(* IEC 61131-3 sources: daoli-st-library/DL_Algo (part 9) *)

(* ---- FB_DL_CascadeCtrl.st ---- *)
(*==============================================================================
 * 组件名称 (Component)  : FB_DL_CascadeCtrl
 * 所属子库 (Sublibrary) : DL_Algo
 * 当前版本 (Version)    : 1.0.0
 * 兼容性   (Platform)   : CODESYS 3.5 / TwinCAT 3 / 汇川 InoProShop / Machine Expert
 *                         仅依赖 Standard.library（R_TRIG），零厂商方言
 * 来源标签 (Source)     : self-std（控制族新增线）
 * 功能描述 (Function)   : 串级控制**骨架**：主回路 PID 输出作从回路外设定，从回路输出
 *                         驱动执行器；双向抗积分饱和（从回路输出饱和时冻结主回路积分）
 *                         + 手动切串级无扰（主 / 从两环积分分别回投跟踪）。
 * 分工互引 (Boundary)   : ① FB_DL_CascadePid 是「双 PID 直连组合件」，只做手动/串级
 *                         两态与副设定钳位；本件是**骨架件**：把抗饱和回投、从环跟踪、
 *                         切换无扰三件事做成显式状态与显式出口，供上层工站编排；
 *                         ② 分程控制归 FB_DL_SplitRangeControl（单回路双阀），与本件
 *                         双回路结构不同；③ 限速归 FB_DL_RateLimiter（本件不做斜坡）。
 * 边界与语义披露 (Boundary disclosure) :
 *   1) 抗饱和口径（条件积分）：从回路输出处于饱和（>= 上限或 <= 下限）且误差同向时，
 *      冻结主回路积分累加（不再朝饱和方向推进）；反向误差照常积分（可自然退出饱和）。
 *   2) 无扰切换：eManual -> eCascade 的切换拍，主回路积分预置为
 *      fSpSlaveLast − fKpM × eM，从回路积分预置为 fManualOut − fKpS × eS，
 *      使切换拍输出连续（验收向量见头注释末行）。
 *   3) 采样时间 tSample 只用于积分折算，fDtSec 由 TIME 转得并参与有限闸（R272）；
 *      tSample <= T#0S 属组态非法。
 *   4) 组态域闸全枚举全部浮点入参（R272）：主/从 PV 与设定、四个增益、四个限值、
 *      fDtSec 全部进入有限性判据；Inf 才是真穿透通道，故不许漏项。
 *   5) 非有限输入：本拍不推进积分（冻结保持上一拍积分量），输出保持上一拍值，
 *      置故障级码并锁存至复位沿 + 输入恢复（污染值绝不允许进入积分器）。
 * 故障码表 (Error codes) :
 *   16#0002_3750 [故障级] 组态非法（限值反向 / 增益非有限 / 采样周期非正）
 *                 反证：冻结保持与「设定恰好等于反馈」输出组合相同，无码不可区分。
 *   16#0002_3751 [故障级] 输入非有限（PV 或设定），积分冻结且输出保持
 *                 反证：保持与「误差为零自然稳态」输出相同，无码则 NaN 事故静默。
 *   16#0002_3753 [信息级] 抗饱和生效（主回路积分被冻结，bAntiWindup 同源可查）
 *                 反证：积分冻结是内部行为，输出上看不出「本拍本该多积多少」。
 * 码位总账 (Code ledger) : 16#0002_3750 / 3751 用 ｜ 16#0002_3753 用
 * 依赖     (Depends)    : 无 DL_ 内部依赖；Standard.library: R_TRIG
 * 红线自检 (Redline)    : R1 ✓ 零全局变量 ｜ R2 ✓ 零 %I/%Q ｜ R3 ✓ 纯 IEC 61131-3
 *                         R4 ✓ 除零闸（fDtSec 由组态闸保证 > 0）/ 非有限三判 / 域闸全枚举
 *                         R5 ✓ 全变量双语同行注释 ｜ R6 ✓ 四态 ENUM + ELSE 兜底
 *                         R7 ✓ 一沿实例主体最前部无条件刷新
 * 修订历史 (Revision)   : 2026-11-22  v1.0.0  首版入库（R69 构建轮 · 批 3 · N9）
 *   验收向量：V1 串级跟随（主设定阶跃 -> 从设定平滑且钳在域内）；V2 抗饱和（从输出
 *             顶到上限时主积分不再增长）；V3 无扰切换（手动 40.0 切串级首拍输出 40.0）；
 *             V4 非有限（PV 写 NaN -> 输出保持 + 3751 锁存，复位沿后恢复）
 *============================================================================*)

(*-----------------------------------------------------------------------------
 * 枚举: E_DL_CascCtrlState（归属 DL_Algo，与 FB_DL_CascadeCtrl 同文件）
 *----------------------------------------------------------------------------*)
TYPE E_DL_CascCtrlState :
(
    eIdle    := 0,    // 未使能：输出下限（安全侧）/ Disabled, output at the lower limit
    eCascade := 10,   // 串级自动：主环驱动从环 / Cascade, master drives the slave
    eManual  := 20,   // 手动：从环手动输出，两环跟踪 / Manual, slave manual, both loops tracking
    eFault   := 99    // 故障锁存：输出保持上一拍 / Fault latched, output holds the last value
);
END_TYPE

(*==============================================================================
 * 功能块: FB_DL_CascadeCtrl
 * 调用约定: 每个扫描周期无条件调用一次。
 *============================================================================*)
FUNCTION_BLOCK FB_DL_CascadeCtrl
VAR_INPUT
    fSpMaster   : REAL := 0.0;              // 主回路设定 [工程单位] / master setpoint
    fPvMaster   : REAL := 0.0;              // 主回路测量 [工程单位] / master process value
    fPvSlave    : REAL := 0.0;              // 从回路测量 [工程单位] / slave process value
    fKpM        : REAL := 1.0;              // 主回路比例增益 [无量纲] / master proportional gain
    fKiM        : REAL := 0.1;              // 主回路积分增益 [1/s] / master integral gain
    fKpS        : REAL := 1.0;              // 从回路比例增益 [无量纲] / slave proportional gain
    fKiS        : REAL := 0.5;              // 从回路积分增益 [1/s] / slave integral gain
    fSpSlaveMin : REAL := 0.0;              // 从回路外设定下限 [工程单位] / slave setpoint floor
    fSpSlaveMax : REAL := 100.0;            // 从回路外设定上限 [工程单位] / slave setpoint ceiling
    fOutMin     : REAL := 0.0;              // 执行器输出下限 [%] / actuator output floor [%]
    fOutMax     : REAL := 100.0;            // 执行器输出上限 [%] / actuator output ceiling [%]
    tSample     : TIME := T#100MS;          // 采样周期 [ms]，<= T#0S 组态非法 / sample period [ms]
    bCascadeMode: BOOL := TRUE;             // TRUE = 串级自动，FALSE = 手动 / TRUE cascade, FALSE manual
    fManualOut  : REAL := 0.0;              // 手动输出 [%] / manual output [%]
    bEnable     : BOOL := TRUE;             // 使能 / enable
    bReset      : BOOL;                     // 上升沿：清故障锁存 / rising edge clears the fault latch
END_VAR
VAR_OUTPUT
    fOut        : REAL;                     // 执行器输出 [%]，域 [fOutMin, fOutMax] / actuator output [%]
    fSpSlave    : REAL;                     // 从回路生效外设定 [工程单位] / effective slave setpoint
    bAntiWindup : BOOL;                     // 抗饱和生效（主积分被冻结）/ anti-windup active
    bSaturated  : BOOL;                     // 从回路输出饱和 / slave output saturated
    bError      : BOOL;                     // 故障标志（组态 / 非有限锁存）/ fault flag
    uErrorId    : UDINT;                    // 故障码，0 = 无故障 / error code, 0 = none
    eState      : E_DL_CascCtrlState;       // 当前状态（供 HMI 诊断）/ current state
END_VAR
VAR
    fbTrigReset : R_TRIG;                   // 复位沿检测实例 / reset edge detector
    eStateInt   : E_DL_CascCtrlState;       // 主状态机内部当前态 / internal state
    eStatePrev  : E_DL_CascCtrlState;       // 上一拍状态（切换沿判据）/ previous state for the transfer edge
    fDtSec      : REAL;                     // 采样周期折算 [s]，参与有限闸 / sample period in seconds, gated
    fErrM       : REAL;                     // 主回路误差 [工程单位] / master error
    fErrS       : REAL;                     // 从回路误差 [工程单位] / slave error
    fIntM       : REAL;                     // 主回路积分累加量 [工程单位] / master integral term
    fIntS       : REAL;                     // 从回路积分累加量 [%] / slave integral term
    fSpSlaveRaw : REAL;                     // 未钳的从回路外设定 [工程单位] / unclamped slave setpoint
    fOutRaw     : REAL;                     // 未钳的执行器输出 [%] / unclamped actuator output
    fOutHold    : REAL;                     // 输出保持值（非有限期）[%] / held output value
    bInBad      : BOOL;                     // 本拍输入非有限 / input non-finite this scan
    bCfgBad     : BOOL;                     // 本拍组态非法 / config illegal this scan
    bCfgLatch   : BOOL;                     // 组态锁存（复位沿 + 组态改对解除）/ config latch
    bFaultLatch : BOOL;                     // 非有限锁存（复位沿 + 输入恢复解除）/ non-finite latch
    bSatInt     : BOOL;                     // 从回路输出饱和内部副本 / internal saturation flag
    bErrorInt   : BOOL;                     // 本拍故障置位累加（出口归并）/ fault set accumulator
    bFirstScan  : BOOL := TRUE;             // 上电首扫标志 / first-scan flag
END_VAR
VAR CONSTANT
    DL_CC_FIN_LIM : REAL := 1.0E30;         // REAL 幅值兜底判界 / REAL magnitude bound
    DL_CC_MS_TO_S : REAL := 1000.0;         // 毫秒到秒折算常数 [ms/s] / milliseconds per second
END_VAR
VAR
    nSampleMs   : DINT;                     // 采样周期整毫秒 [ms] / sample period in whole milliseconds
END_VAR

(*------------------------------------------------------------------------------
 * 段 1｜无条件刷新区（红线 R7）：一沿实例位于主体最前部
 *      Unconditional refresh: the edge instance at the very top
 *-----------------------------------------------------------------------------*)
fbTrigReset(CLK := bReset);

(* 段 2｜上电首扫：积分与输出落安全侧 / first-scan init *)
IF bFirstScan THEN
    eStateInt  := E_DL_CascCtrlState.eIdle;
    eStatePrev := E_DL_CascCtrlState.eIdle;
    fIntM      := 0.0;
    fIntS      := 0.0;
    fOutHold   := 0.0;
    bFirstScan := FALSE;
END_IF

(* 段 3｜每拍预清（FB32-1）：单拍标志，禁入积分 / per-scan preset *)
bSatInt := FALSE;

bErrorInt := FALSE;                     // 每拍预清（单拍标志）/ per-scan preset

(*------------------------------------------------------------------------------
 * 段 4｜组态域闸（R151 / R272 全枚举）：四个限值序 + 四个增益 + 采样周期 + fDtSec
 *      Config gate over the limits, the gains, the sample period and fDtSec
 *      解除路径（R152 自证可达）：复位沿 AND 组态非法条件全部消失
 *-----------------------------------------------------------------------------*)
nSampleMs := TIME_TO_DINT(tSample);     // TIME -> 整毫秒（标准转换函数）/ TIME to milliseconds
fDtSec    := DINT_TO_REAL(nSampleMs) / DL_CC_MS_TO_S;   // 毫秒 -> 秒（除子为常数 1000 > 0）[s] / to seconds

bCfgBad := (fSpSlaveMin >= fSpSlaveMax) OR (fOutMin >= fOutMax)
           OR (fSpSlaveMin <> fSpSlaveMin) OR (fSpSlaveMax <> fSpSlaveMax)
           OR (fOutMin <> fOutMin) OR (fOutMax <> fOutMax)
           OR (fKpM <> fKpM) OR (fKiM <> fKiM) OR (fKpS <> fKpS) OR (fKiS <> fKiS)
           OR (ABS(fKpM) >= DL_CC_FIN_LIM) OR (ABS(fKiM) >= DL_CC_FIN_LIM)
           OR (ABS(fKpS) >= DL_CC_FIN_LIM) OR (ABS(fKiS) >= DL_CC_FIN_LIM)
           OR (ABS(fSpSlaveMin) >= DL_CC_FIN_LIM) OR (ABS(fSpSlaveMax) >= DL_CC_FIN_LIM)
           OR (ABS(fOutMin) >= DL_CC_FIN_LIM) OR (ABS(fOutMax) >= DL_CC_FIN_LIM)
           OR (tSample <= T#0S) OR (fDtSec <= 0.0) OR (fDtSec <> fDtSec)
           OR (ABS(fDtSec) >= DL_CC_FIN_LIM);

IF bCfgBad THEN
    bCfgLatch := TRUE;
END_IF
IF fbTrigReset.Q AND (NOT bCfgBad) THEN
    bCfgLatch := FALSE;                   // 组态锁存解除 / config latch cleared
    uErrorId  := 16#0000_0000;            // 码位随解除归零 / code cleared with the latch
END_IF
IF bCfgLatch THEN
    uErrorId  := 16#0002_3750;            // 故障级：组态非法 / fault: illegal configuration
    bErrorInt := TRUE;                    // R45 配对 / paired with the code
    eStateInt := E_DL_CascCtrlState.eFault;
END_IF

(*------------------------------------------------------------------------------
 * 段 5｜输入有限闸（R272）：PV 与设定全部入闸；非有限即锁存并冻结积分
 *      Input finiteness gate: any non-finite PV freezes the integrals and holds the output
 *-----------------------------------------------------------------------------*)
bInBad := (fSpMaster <> fSpMaster) OR (fPvMaster <> fPvMaster) OR (fPvSlave <> fPvSlave)
          OR (fManualOut <> fManualOut)
          OR ((fSpMaster - fSpMaster) <> (fSpMaster - fSpMaster))
          OR ((fPvMaster - fPvMaster) <> (fPvMaster - fPvMaster))
          OR ((fPvSlave - fPvSlave) <> (fPvSlave - fPvSlave))
          OR (ABS(fSpMaster) >= DL_CC_FIN_LIM) OR (ABS(fPvMaster) >= DL_CC_FIN_LIM)
          OR (ABS(fPvSlave) >= DL_CC_FIN_LIM) OR (ABS(fManualOut) >= DL_CC_FIN_LIM);

IF bInBad THEN
    bFaultLatch := TRUE;
END_IF
IF fbTrigReset.Q AND (NOT bInBad) THEN
    bFaultLatch := FALSE;                 // 非有限锁存解除（复位沿 + 输入恢复）/ latch cleared once the input is finite
    uErrorId    := 16#0000_0000;
END_IF

(*------------------------------------------------------------------------------
 * 段 6｜主状态机（红线 R6）：ENUM + CASE + ELSE 兜底
 *      Main state machine, phase semantics only
 *-----------------------------------------------------------------------------*)
CASE eStateInt OF

    E_DL_CascCtrlState.eIdle:
        IF bEnable AND (NOT bCfgLatch) AND (NOT bFaultLatch) THEN
            IF bCascadeMode THEN
                eStateInt := E_DL_CascCtrlState.eCascade;
            ELSE
                eStateInt := E_DL_CascCtrlState.eManual;
            END_IF
        END_IF

    E_DL_CascCtrlState.eCascade:
        IF (NOT bEnable) OR bCfgLatch OR bFaultLatch THEN
            eStateInt := E_DL_CascCtrlState.eIdle;
        ELSIF NOT bCascadeMode THEN
            eStateInt := E_DL_CascCtrlState.eManual;    // 切手动（从环手动，主环跟踪）/ to manual with tracking
        END_IF

    E_DL_CascCtrlState.eManual:
        IF (NOT bEnable) OR bCfgLatch OR bFaultLatch THEN
            eStateInt := E_DL_CascCtrlState.eIdle;
        ELSIF bCascadeMode THEN
            eStateInt := E_DL_CascCtrlState.eCascade;   // 切串级（切换拍做无扰回投）/ to cascade with bumpless transfer
        END_IF

    E_DL_CascCtrlState.eFault:
        IF fbTrigReset.Q AND (NOT bCfgBad) AND (NOT bInBad) THEN
            bCfgLatch := FALSE;                         // 两类锁存同沿解除 / both latches cleared together
            bFaultLatch := FALSE;
            uErrorId  := 16#0000_0000;
            eStateInt := E_DL_CascCtrlState.eIdle;
        END_IF

    ELSE
        (* 非法状态拦截 / illegal state interception *)
        eStateInt := E_DL_CascCtrlState.eFault;
        uErrorId  := 16#0002_3750;
        bErrorInt := TRUE;

END_CASE;

(*------------------------------------------------------------------------------
 * 段 7｜主 / 从两环求值与抗饱和回投（条件积分口径）
 *      Master and slave evaluation with conditional-integration anti-windup
 *-----------------------------------------------------------------------------*)
fErrM := fSpMaster - fPvMaster;                 // 主回路误差 [工程单位] / master error
fErrS := 0.0;                                   // 从回路误差缺省 0（从设定在下段算出）/ slave error default
bAntiWindup := FALSE;

IF (NOT bInBad) AND (NOT bCfgLatch) AND (eStateInt <> E_DL_CascCtrlState.eFault) THEN
    IF eStateInt = E_DL_CascCtrlState.eManual THEN
        (* 手动：从环手动输出，两环做跟踪回投（直接零跳变）/ manual with loop tracking *)
        fIntS := fManualOut - fKpS * (fSpSlave - fPvSlave);   // 从环积分回投 [%] / slave integral back-injected
        fIntM := fSpSlave - fKpM * fErrM;                     // 主环积分回投（输出即从设定）[工程单位] / master integral back-injected
    ELSE
        (* 串级：主环条件积分（从环饱和且误差同向时冻结）/ cascade with conditional integration *)
        IF bSatInt AND (((fSpSlave >= fSpSlaveMax) AND (fErrM > 0.0)) OR ((fSpSlave <= fSpSlaveMin) AND (fErrM < 0.0))) THEN
            bAntiWindup := TRUE;                   // 冻结主积分（不再朝饱和方向推进）/ freeze the master integral
            uErrorId    := 16#0002_3753;           // 信息级：抗饱和生效 / info: anti-windup active
        ELSE
            fIntM := fIntM + fKiM * fErrM * fDtSec;   // 主积分推进 [工程单位] / master integral step
        END_IF
        fSpSlaveRaw := fKpM * fErrM + fIntM;       // 主环输出即从环设定 [工程单位] / master output is the slave setpoint
        IF fSpSlaveRaw > fSpSlaveMax THEN
            fSpSlaveRaw := fSpSlaveMax;            // 从设定钳上限 / clamp the slave setpoint
        ELSIF fSpSlaveRaw < fSpSlaveMin THEN
            fSpSlaveRaw := fSpSlaveMin;            // 从设定钳下限 / clamp the slave setpoint
        END_IF
        fErrS := fSpSlaveRaw - fPvSlave;           // 从回路误差 [工程单位] / slave error
        fIntS := fIntS + fKiS * fErrS * fDtSec;    // 从积分推进 [%] / slave integral step
    END_IF
END_IF

(*------------------------------------------------------------------------------
 * 段 8｜输出合成与限幅（非有限期保持上一拍值）/ output folding with the hold path
 *-----------------------------------------------------------------------------*)
IF (eStateInt = E_DL_CascCtrlState.eManual) THEN
    fOutRaw := fManualOut;                         // 手动：直出手动值 [%] / manual pass-through
ELSE
    fOutRaw := fKpS * fErrS + fIntS;               // 串级：从环 PI 输出 [%] / slave PI output
END_IF

IF fOutRaw > fOutMax THEN
    fOutRaw  := fOutMax;                           // 输出钳上限 [%] / clamp high
    bSatInt  := TRUE;
ELSIF fOutRaw < fOutMin THEN
    fOutRaw  := fOutMin;                           // 输出钳下限 [%] / clamp low
    bSatInt  := TRUE;
END_IF

IF bInBad OR bCfgLatch THEN
    fOut := fOutHold;                              // 非有限 / 组态故障：保持上一拍（不注入污染值）[%] / hold
    IF bInBad THEN
        uErrorId  := 16#0002_3751;                 // 故障级：输入非有限 / fault: non-finite input
        bErrorInt := TRUE;                         // R45 配对 / paired with the code
    END_IF
ELSIF eStateInt = E_DL_CascCtrlState.eIdle THEN
    fOut := fOutMin;                               // 未使能：输出下限（安全侧）[%] / disabled, output floor
ELSE
    fOut := fOutRaw;                               // 正常：限幅后输出 [%] / normal path
END_IF
fOutHold := fOut;                                  // 保持值快照（主体末行）/ snapshot the hold value

(*------------------------------------------------------------------------------
 * 段 9｜输出单一出口（范式 P-05）
 *      Single output exit
 *-----------------------------------------------------------------------------*)
IF eStateInt = E_DL_CascCtrlState.eCascade THEN
    fSpSlave := fSpSlaveRaw;                       // 串级：生效从设定即主环输出 [工程单位] / effective slave setpoint
ELSE
    fSpSlave := fPvSlave;                          // 手动 / 空闲：从设定跟实测（跟踪位置）[工程单位] / tracking position
END_IF
bSaturated := bSatInt;
bError     := bErrorInt OR bCfgLatch OR bFaultLatch;
eState     := eStateInt;
eStatePrev := eStateInt;                           // 状态快照刷新（供下一拍切换沿判据）/ refresh the state snapshot
END_FUNCTION_BLOCK

(* ---- FB_DL_CascadePid.st ---- *)
(*==============================================================================
 * 组件名称 (Component)  : FB_DL_CascadePid
 * 所属子库 (Sublibrary) : DL_Algo
 * 当前版本 (Version)    : 1.0.0
 * 兼容性   (Platform)   : CODESYS 3.5 / TwinCAT 3 / 汇川 InoProShop / Machine Expert
 *                         仅依赖 Standard.library（R_TRIG 间接经子块），零厂商方言
 * 功能描述 (Function)   : 主副双回路串级 PID。主回路 PID 输出经限幅后作为副回路
 *                         设定值，副回路输出驱动执行器；适用温控（主温度 / 副加
 *                         热功率）、张力（主张力 / 副速度）等场景。内部组合两个
 *                         FB_DL_PidController 实例，本块不自写 PID 律；手动时副
 *                         回路直接手动输出，主回路经跟踪回投跟随副设定，回自动
 *                         零跳变。两个实例的采样周期与输出限幅统一由本块注入，
 *                         杜绝调用方双份配置不一致。
 * 开源溯源 (Origin)     : 原创实现。串级结构分类与参数域参考 OSCAT / 西门子
 *                         CASCADE_CONT 的公开语义描述，未复制任何厂商源码。
 * 本文件内含       : TYPE  E_DL_CascadeState（配套枚举，归属 DL_Algo）
 *                    FB    FB_DL_CascadePid
 * 依赖     (Depends)    : FB_DL_PidController（DL_Algo 内部）
 * 红线自检 (Redline)    : R1 ✓ 零全局变量表与外部变量引用 ｜ R2 ✓ 零物理 IO 地址直写
 *                         R3 ✓ 纯 IEC 61131-3 ｜ R4 ✓ 防除零+钳位+非有限值防御
 *                         R5 ✓ 全变量中英双语同行注释 ｜ R6 ✓ 四态 ENUM+CASE+ELSE
 *                         R7 ✓ 定时器 / 边沿实例均由子块无条件刷新（本块无实例）
 * 修订历史 (Revision)   :
 *   2026-11-15  v1.0.0  首版入库 · Round 04 · Level 1 DL_Algo
 * 验收向量 (Acceptance) :
 *   V1 串级跟随：主设定阶跃 50 → fSpSlave 平滑爬升并钳在副设定域内
 *   V2 副设定钳位：主回路输出超 rSpSlaveMax → fSpSlave 恰等于 rSpSlaveMax
 *   V3 手动无扰：手动副输出 40.0 切串级首拍 fOut 保持 40.0 连续
 *   V4 参数对调：rSpSlaveMin>rSpSlaveMax 时自动对调且 uErrorId=0002_0001
 *   V5 非有限值：fPvSlave 写入非法浮点 → 输出保持上一拍且 uErrorId=0002_0004
 *============================================================================*)

(*-----------------------------------------------------------------------------
 * 枚举: E_DL_CascadeState（归属 DL_Algo，与 FB_DL_CascadePid 同文件）
 * 含义: 串级控制器离散状态。数值步长留空位便于后续插态而不破坏已有工程。
 *----------------------------------------------------------------------------*)
TYPE E_DL_CascadeState :
(
    eIdle    := 0,    // 使能关：双回路冻结，输出回下限 / Idle: enable off, both loops frozen
    eCascade := 10,   // 双回路自动：主环驱动副环闭环 / Cascade: master drives slave in closed loop
    eManual  := 20,   // 手动：副环手动输出，主环跟踪副设定 / Manual: slave manual, master tracks slave SP
    eFault   := 99    // 故障兜底态：非法状态进入，输出安全值 / Fault fallback: illegal state, safe output
);
END_TYPE

(*==============================================================================
 * 功能块: FB_DL_CascadePid
 * 调用约定: 每个扫描周期无条件调用一次；bReset 电平透传给两个子块。
 * 无状态泄漏: 全部状态驻留于实例私有 VAR，零全局引用，可多实例并行。
 * 架构披露: 本块零自写 PID 律，仅做设定值路由、限幅注入与状态调度。
 *============================================================================*)
FUNCTION_BLOCK FB_DL_CascadePid
VAR_INPUT
    bEnable          : BOOL := FALSE;   // 总使能，FALSE 时输出回下限 / Master enable, FALSE drives output to low limit
    bManual          : BOOL := FALSE;   // 手动模式，TRUE 时副环手动 / Manual mode, TRUE puts slave loop in manual
    fManualSlaveValue: REAL := 0.0;     // 副回路手动输出 [%] / Slave loop manual output in percent
    fSpMaster        : REAL := 0.0;     // 主回路设定值 [EU] / Master loop setpoint in engineering units
    fPvMaster        : REAL := 0.0;     // 主回路过程值 [EU] / Master loop process value
    fPvSlave         : REAL := 0.0;     // 副回路过程值 [EU] / Slave loop process value
    fKpM             : REAL := 1.0;     // 主回路比例增益 [1] / Master loop proportional gain
    tTiM             : TIME := T#5S;    // 主回路积分时间 [s] / Master loop integral time
    tTdM             : TIME := T#0S;    // 主回路微分时间 [s] / Master loop derivative time
    fKpS             : REAL := 2.0;     // 副回路比例增益 [1]，默认更硬 / Slave gain, harder by default
    tTiS             : TIME := T#1S;    // 副回路积分时间 [s] / Slave loop integral time
    tTdS             : TIME := T#0S;    // 副回路微分时间 [s] / Slave loop derivative time
    rSpSlaveMin      : REAL := 0.0;     // 副设定域下限 [EU] / Slave setpoint domain lower limit
    rSpSlaveMax      : REAL := 100.0;   // 副设定域上限 [EU] / Slave setpoint domain upper limit
    rOutMin          : REAL := 0.0;     // 副环输出下限 [%] / Slave output lower limit in percent
    rOutMax          : REAL := 100.0;   // 副环输出上限 [%] / Slave output upper limit in percent
    tSampleTime      : TIME := T#100MS; // 采样周期，统一注入两个子块 / Sample period injected to both sub-blocks
    bReset           : BOOL := FALSE;   // 复位信号，电平透传两个子块 / Reset passed through to both sub-blocks
END_VAR
VAR_OUTPUT
    fOut             : REAL;            // 副回路控制输出 [%] / Slave loop control output in percent
    fSpSlave         : REAL;            // 副回路设定值 [EU]，诊断 / Slave setpoint in engineering units, diagnostics
    fErrMaster       : REAL;            // 主回路偏差 [EU]，诊断 / Master loop error, diagnostics
    bLimitHigh       : BOOL;            // 副环输出触上限 / Slave output at upper limit
    bLimitLow        : BOOL;            // 副环输出触下限 / Slave output at lower limit
    bError           : BOOL;            // 故障标志 / Fault flag
    uErrorId         : UDINT;           // 故障码，0 = 无故障 / Error code, 0 = no error
END_VAR
VAR
    fbPidMaster      : FB_DL_PidController;  // 主回路 PID 实例 / Master loop PID instance
    fbPidSlave       : FB_DL_PidController;  // 副回路 PID 实例 / Slave loop PID instance
    eState           : E_DL_CascadeState;    // 主状态机当前状态 / Current state of the state machine
    fSpSlaveLow      : REAL;            // 对调修复后的副设定域下限 [EU] / Repaired slave SP domain low limit
    fSpSlaveHigh     : REAL;            // 对调修复后的副设定域上限 [EU] / Repaired slave SP domain high limit
    fMasterOutClamp  : REAL;            // 钳位到副设定域的主回路输出 [EU] / Master output clamped into slave domain
    bNonFinite       : BOOL;            // 本拍输入非有限值标志 / Non-finite input flag of this cycle
END_VAR

(*------------------------------------------------------------------------------
 * 段 1｜参数钳位与公共防御（不中断扫描）
 *      Parameter clamping and common defenses, never stops the scan
 *-----------------------------------------------------------------------------*)
bError   := FALSE;                    // 每拍重算故障标志 / Recompute fault flag every cycle
uErrorId := 16#0002_0000;             // 每拍重算故障码 / Recompute error code every cycle
bLimitHigh := FALSE;                  // 触限标志每拍重算 / Saturation flags recomputed every cycle
bLimitLow  := FALSE;                  // 触限标志每拍重算 / Saturation flags recomputed every cycle
bNonFinite := FALSE;                  // 非有限值标志每拍重算 / Non-finite flag recomputed every cycle

IF tSampleTime < T#10MS THEN
    tSampleTime := T#10MS;            // 采样周期非法钳位为 10 ms / Illegal sample period clamped to 10 ms
    uErrorId := 16#0002_0002;         // 公共码：采样周期已钳位 / Common code: sample period clamped
END_IF

IF rSpSlaveMin > rSpSlaveMax THEN
    fSpSlaveLow  := rSpSlaveMax;      // 对调修复（下限取原上限） / Swapped repair of domain low limit
    fSpSlaveHigh := rSpSlaveMin;      // 对调修复（上限取原下限） / Swapped repair of domain high limit
    uErrorId := 16#0002_0001;         // 公共码：参数越界已钳位 / Common code: parameter clamped
ELSE
    fSpSlaveLow  := rSpSlaveMin;      // 合法域下限直通 / Valid domain low limit passed
    fSpSlaveHigh := rSpSlaveMax;      // 合法域上限直通 / Valid domain high limit passed
END_IF

(* 输入非有限值防御：任一主 / 副回路信号非法即拒绝本拍更新 *)
(* Non-finite defense: reject this cycle if any master or slave signal invalid *)
IF (fSpMaster <> fSpMaster) OR (ABS(fSpMaster) > 1.0E30)
   OR (fPvMaster <> fPvMaster) OR (ABS(fPvMaster) > 1.0E30)
   OR (fPvSlave <> fPvSlave) OR (ABS(fPvSlave) > 1.0E30)
   OR (fManualSlaveValue <> fManualSlaveValue) OR (ABS(fManualSlaveValue) > 1.0E30) THEN
    bNonFinite := TRUE;               // 置非有限值标志 / Set non-finite flag
END_IF

(*------------------------------------------------------------------------------
 * 段 2｜子块统一注入：两个实例的采样周期与输出限幅由本块独占配置
 *      Unified injection: sample period and output limits owned by this block
 *-----------------------------------------------------------------------------*)
fbPidMaster.bEnable     := bEnable AND (NOT bManual) AND (NOT bNonFinite);
fbPidMaster.fSetpoint   := fSpMaster;             // 主设定注入 / Inject master setpoint
fbPidMaster.fActual     := fPvMaster;             // 主过程值注入 / Inject master process value
fbPidMaster.fKp         := fKpM;                  // 主增益注入 / Inject master gain
fbPidMaster.tTi         := tTiM;                  // 主积分时间注入 / Inject master integral time
fbPidMaster.tTd         := tTdM;                  // 主微分时间注入 / Inject master derivative time
fbPidMaster.fDeadband   := 0.0;                   // 主环死区默认关闭 / Master deadband off by default
fbPidMaster.bIncremental:= FALSE;                 // 主环默认位置式 / Master positional by default
fbPidMaster.rOutMin     := fSpSlaveLow;           // 主输出域 = 副设定域（下限） / Master domain equals slave SP domain
fbPidMaster.rOutMax     := fSpSlaveHigh;          // 主输出域 = 副设定域（上限） / Master domain equals slave SP domain
fbPidMaster.tSampleTime := tSampleTime;           // 统一采样周期 / Unified sample period
fbPidMaster.bTrack      := FALSE;                 // 跟踪在状态机内按需置位 / Tracking set inside state machine
fbPidMaster.fTrackValue := fSpSlave;              // 跟踪值 = 当前副设定 / Track value equals current slave SP
fbPidMaster.bReset      := bReset;                // 复位透传 / Reset passed through

fbPidSlave.bEnable      := bEnable AND (NOT bNonFinite);
fbPidSlave.fSetpoint    := fSpSlave;              // 副设定注入 / Inject slave setpoint
fbPidSlave.fActual      := fPvSlave;              // 副过程值注入 / Inject slave process value
fbPidSlave.fKp          := fKpS;                  // 副增益注入 / Inject slave gain
fbPidSlave.tTi          := tTiS;                  // 副积分时间注入 / Inject slave integral time
fbPidSlave.tTd          := tTdS;                  // 副微分时间注入 / Inject slave derivative time
fbPidSlave.fDeadband    := 0.0;                   // 副环死区默认关闭 / Slave deadband off by default
fbPidSlave.bIncremental := FALSE;                 // 副环默认位置式 / Slave positional by default
fbPidSlave.rOutMin      := rOutMin;               // 副环输出下限注入 / Inject slave output low limit
fbPidSlave.rOutMax      := rOutMax;               // 副环输出上限注入 / Inject slave output high limit
fbPidSlave.tSampleTime  := tSampleTime;           // 统一采样周期 / Unified sample period
fbPidSlave.bTrack       := FALSE;                 // 副环不需要跟踪 / Slave needs no tracking
fbPidSlave.fTrackValue  := 0.0;                   // 跟踪值占位为 0 / Track value placeholder zero
fbPidSlave.bReset       := bReset;                // 复位透传 / Reset passed through

(*------------------------------------------------------------------------------
 * 段 3｜主状态机（红线 R6）：ENUM + CASE + ELSE 兜底
 *      Main state machine: ENUM + CASE with mandatory ELSE fallback
 *-----------------------------------------------------------------------------*)
CASE eState OF

    eIdle:
        (* 使能关：双回路冻结，输出回下限，副设定保持在域下限 *)
        (* Enable off: both loops frozen, output at low limit, slave SP at domain low *)
        fOut       := rOutMin;        // 输出回下限 / Output to low limit
        fSpSlave   := fSpSlaveLow;    // 副设定保持域下限 / Slave SP held at domain low
        fErrMaster := fSpMaster - fPvMaster;  // 主偏差仍刷新供诊断 / Master error for diagnostics
        IF bEnable AND (NOT bNonFinite) THEN
            IF bManual THEN
                eState := eManual;        // 请求手动 / Request manual mode
            ELSE
                eState := eCascade;       // 请求串级自动 / Request cascade auto
            END_IF
        END_IF

    eCascade:
        (* 串级自动：主回路闭环 → 主输出钳位到副设定域 → 副回路闭环 *)
        (* Cascade auto: master closed loop, output clamped into slave domain, slave loop *)
        IF bNonFinite THEN
            (* 非有限值拍：保持上一拍输出，置公共拒绝码 *)
            (* Non-finite cycle: hold previous output, common reject code *)
            bError   := TRUE;             // 置故障标志 / Set fault flag
            uErrorId := 16#0002_0004;     // 输入非有限值已拒绝 / Non-finite input rejected
        ELSE
            fbPidMaster.bEnable := TRUE;  // 主环使能 / Enable master loop
            fbPidMaster();                // 主回路运算 / Master loop computation
            fMasterOutClamp := LIMIT(fSpSlaveLow, fbPidMaster.fOut, fSpSlaveHigh);  // 钳位 / Clamp into slave domain
            IF fbPidMaster.bLimitHigh OR fbPidMaster.bLimitLow THEN
                IF uErrorId = 16#0002_0000 THEN
                    uErrorId := 16#0002_0201;  // 信息级：副设定超域已钳位 / Info: slave SP clamped
                END_IF
            END_IF
            fSpSlave := fMasterOutClamp;  // 副设定 = 钳位后的主输出 / Slave SP equals clamped master output
            fbPidSlave.bEnable := TRUE;   // 副环使能 / Enable slave loop
            fbPidSlave();                 // 副回路运算 / Slave loop computation
            fOut        := fbPidSlave.fOut;       // 输出 = 副环输出 / Output equals slave output
            fErrMaster  := fbPidMaster.fErr;      // 主偏差诊断 / Master error diagnostics
            bLimitHigh  := fbPidSlave.bLimitHigh; // 触限透传 / Saturation passthrough
            bLimitLow   := fbPidSlave.bLimitLow;  // 触限透传 / Saturation passthrough
        END_IF
        IF bManual THEN
            eState := eManual;            // 切手动 / Switch to manual
        ELSIF NOT bEnable THEN
            eState := eIdle;              // 切空闲 / Switch to idle
        END_IF

    eManual:
        (* 手动：副环直接手动输出，主环经跟踪回投跟随副设定，回自动无跳变 *)
        (* Manual: slave manual output, master tracks slave SP for bumpless return *)
        IF bNonFinite THEN
            bError   := TRUE;             // 置故障标志 / Set fault flag
            uErrorId := 16#0002_0004;     // 输入非有限值已拒绝 / Non-finite input rejected
        ELSE
            fbPidSlave.bEnable    := TRUE;             // 副环使能 / Enable slave loop
            fbPidSlave.bManual    := TRUE;             // 副环手动 / Slave in manual
            fbPidSlave.fManualValue := fManualSlaveValue;  // 手动值注入 / Inject manual value
            fbPidSlave();                              // 副环手动运算 / Slave manual computation
            fbPidSlave.bManual    := FALSE;            // 恢复自动配置位 / Restore auto config bit
            fOut       := fbPidSlave.fOut;             // 输出 = 副环手动值 / Output equals slave manual value
            fSpSlave   := fSpSlaveLow;                 // 副设定保持在域下限 / Slave SP held at domain low
            fbPidMaster.bEnable    := TRUE;            // 主环使能 / Enable master loop
            fbPidMaster.bManual    := TRUE;            // 主环手动跟踪模式 / Master in manual-track mode
            fbPidMaster.fManualValue := fSpSlaveLow;   // 手动值取域下限占位 / Manual value placeholder
            fbPidMaster.bTrack     := TRUE;            // 跟踪回投使能 / Track enable
            fbPidMaster.fTrackValue:= fSpSlaveLow;     // 主环跟随域下限防积分漂移 / Master tracks domain low
            fbPidMaster();                             // 主环跟踪运算 / Master tracking computation
            fbPidMaster.bManual    := FALSE;           // 恢复自动配置位 / Restore auto config bit
            fbPidMaster.bTrack     := FALSE;           // 清跟踪位 / Clear track bit
            fErrMaster := fbPidMaster.fErr;            // 主偏差诊断 / Master error diagnostics
            bLimitHigh  := fbPidSlave.bLimitHigh;      // 触限透传 / Saturation passthrough
            bLimitLow   := fbPidSlave.bLimitLow;       // 触限透传 / Saturation passthrough
        END_IF
        IF NOT bEnable THEN
            eState := eIdle;              // 切空闲 / Switch to idle
        ELSIF NOT bManual THEN
            eState := eCascade;           // 切串级 / Switch to cascade
        END_IF

    eFault:
        (* 故障兜底态：输出安全下限，等待复位解除 *)
        (* Fault fallback: safe low-limit output, released by reset *)
        fOut := rOutMin;                  // 安全输出 / Safe output

    ELSE
        (* 非法状态拦截：任何未定义状态一律进故障兜底，不做隐式恢复 *)
        (* Illegal state interception: any undefined state goes to fault fallback *)
        eState   := eFault;               // 进故障态 / Enter fault state
        bError   := TRUE;                 // 置故障标志 / Set fault flag
        uErrorId := 16#0002_0005;         // 非法状态兜底码 / Illegal state fallback code
        fOut     := rOutMin;              // 安全输出 / Safe output
END_CASE;

(* 子块故障聚合：优先透传副环故障码，无副环故障时透传主环故障码 *)
(* Sub-block fault aggregation: slave code first, then master code *)
IF (NOT bError) AND (uErrorId = 16#0002_0000) THEN
    IF fbPidSlave.bError THEN
        bError   := TRUE;                 // 副环故障置位 / Slave fault set
        uErrorId := fbPidSlave.uErrorId;  // 透传副环故障码 / Pass slave error code
    ELSIF fbPidMaster.bError THEN
        bError   := TRUE;                 // 主环故障置位 / Master fault set
        uErrorId := fbPidMaster.uErrorId; // 透传主环故障码 / Pass master error code
    END_IF
END_IF
END_FUNCTION_BLOCK

(* ---- FB_DL_CascadeWindupLink.st ---- *)
(*
  FB_DL_CascadeWindupLink  —  串级外环→内环设定传递抗饱和联动 / Cascade windup link between outer and inner PID loops
  分类 Category : DL_Algo
  版本 Version  : 1.0.1
  来源 Source   : t2-5-modpid — 串级抗饱和族零检索深化
  溯源 Origin   : clean-room 实现，未复制任何源码行
  功能 Function : 1) 引用 FB_DL_PidController 引脚契约（不改其对外接口）：外环限幅镜像
                  内环限幅（fbOuter.rOutMin/rOutMax := fInnerMin/fInnerMax）；
                  2) 内环饱和（bLimitHigh/bLimitLow 任一）持续 tSatTo → 故障级 03AC/03AD
                  独立锁存（R190 归因唯一）；饱和期间外环经跟踪机制冻结积分：
                  fbOuter.bTrack := TRUE 且 fTrackValue := fbOuter.fOut（保持当前输出）；
                  3) R242 跟踪相退化推演：镜像钳制与冻结仅在 bTrack=FALSE 相生效——
                  调用方外部跟踪 bExtTrack=TRUE 期间，冻结请求让位（信息级 0494），
                  外部跟踪值直通；
                  4) 外环输出非有限 → 03AE 防御兜底锁存。
  返修记录 Rework  :
    2026-11-19  v1.0.1  R42 P0-3 中等返修：v1.0.0 故障相（段 7 故障分支）仅强制
                        bFreeze/bMirror 出口 FALSE，fbOuter.bTrack 残留 TRUE 且
                        fTrackValue 停更——跟踪标志与外环输出钳制名实不一，
                        外环静默冻结积分（P0 派单缺陷③，R191 名实双出口违反）。
                        修复要点：故障分支显式写 fbOuter.bTrack := FALSE
                        （跟踪释放，钳制语义与标志同拍同步），PID 回自主积分
                        由其自身安全侧承载；对外接口签名不变。
  边界 Boundary : ① 组态闸：fInnerMax <= fInnerMin → 03AB 锁存，镜像与冻结全部停发；
                  ② fbOuter 为 VAR_IN_OUT 引用：写其 rOutMin/rOutMax/bTrack/fTrackValue，
                  读其 fOut/bLimitHigh/bLimitLow/bLimitLow——不改 PidController 对外契约；
                  ③ 解除式全当拍量（R240 落地），逐 BOOL 标注见段 4；
                  ④ 无 GVL 依赖：纯引脚输入输出，无外部变量引用，无物理 IO 地址。
  依赖 Depends  : FB_DL_PidController（注入，不实例化，引脚按 registry 实名）；Standard.library（TON / R_TRIG）
  码表 Error codes（Algo 段 0002，窗口 03AB~03AE / 0491~0494）:
    16#0002_03AB 故障级：组态非法（内环限幅上下界颠倒），锁存至 bReset
    16#0002_03AC 故障级：内环上饱和持续（tSatTo），锁存至 bReset
    16#0002_03AD 故障级：内环下饱和持续（tSatTo），锁存至 bReset
    16#0002_03AE 故障级：外环输出非有限（防御兜底），锁存至 bReset
    16#0002_0491 信息级：镜像钳制生效沿（限幅镜像首次写入）
    16#0002_0492 信息级：外环积分冻结激活沿
    16#0002_0493 信息级：冻结解除恢复沿
    16#0002_0494 信息级：外部跟踪让位（bExtTrack 期间冻结请求被让位）
  修订历史 Revision :
    2026-11-19  v1.0.0  R41 首版（批次 3 · 序号 5）
    2026-11-19  v1.0.1  R42 P0-3 中等返修（见返修记录节）
*)

FUNCTION_BLOCK FB_DL_CascadeWindupLink
VAR_INPUT
    fInnerMin    : REAL := 0.0;       // 内环限幅下限 [%]，必须 < fInnerMax / Inner loop lower limit
    fInnerMax    : REAL := 100.0;     // 内环限幅上限 [%]，必须 > fInnerMin / Inner loop upper limit
    tSatTo       : TIME := T#1S;      // 饱和确认超时 [ms]，域 > 0 / Saturation confirm timeout
    bExtTrack    : BOOL := FALSE;     // 调用方外部跟踪请求 [-] / External tracking request from caller
    fExtTrackVal : REAL := 0.0;       // 外部跟踪值 [%] / External track value
    bEnable      : BOOL := FALSE;     // 联动使能 [-] / Link enable
    bReset       : BOOL := FALSE;     // 复位，上升沿清故障锁存 / Reset edge clears fault latch
END_VAR
VAR_IN_OUT
    fbOuter      : FB_DL_PidController;   // 外环 PID 引用（镜像钳制目标）/ Outer loop PID reference
    fbInner      : FB_DL_PidController;   // 内环 PID 引用（饱和判据来源）/ Inner loop PID reference
END_VAR
VAR_OUTPUT
    bFreeze      : BOOL;              // 外环冻结标志（实际生效）[-] / Effective freeze flag
    bMirror      : BOOL;              // 限幅镜像生效标志 [-] / Mirror active flag
    bError       : BOOL;              // 故障锁存标志 / Fault latch flag
    nErrId       : UDINT;             // 事件码，0 = 无事件 / Event code
END_VAR
VAR
    tonSatHiTo   : TON;               // 上饱和确认定时器（专用超时命名），无条件刷新 / High-saturation timer
    tonSatLoTo   : TON;               // 下饱和确认定时器（专用超时命名），无条件刷新 / Low-saturation timer
    rtReset      : R_TRIG;            // 复位沿实例，无条件刷新 / Reset edge instance
    _bSatHigh    : BOOL;              // 内环上饱和当拍量 [-] / Inner high-saturation flag
    _bSatLow     : BOOL;              // 内环下饱和当拍量 [-] / Inner low-saturation flag
    _bHiLat      : BOOL;              // 上饱和锁存位（锁存量）/ High-saturation latch bit
    _bLoLat      : BOOL;              // 下饱和锁存位（锁存量）/ Low-saturation latch bit
    _bCfgBad     : BOOL;              // 组态锁存位（锁存量）/ Config-fault latch bit
    _uFault      : UDINT;             // 故障码锁存（锁存量）/ Latched fault code
    _uInfo       : UDINT;             // 信息码，每拍重算 / Transient info code
    _bMirrorSent : BOOL;              // 镜像首次写入沿判据快照 / Mirror first-write edge snapshot
    _bFreezePrev : BOOL;              // 上拍冻结镜像（解除沿判据）/ Previous freeze mirror
END_VAR

(* —— 段 0：定时器与沿实例无条件周期刷新（禁置于 IF/CASE 内） —— *)
_bSatHigh := fbInner.bLimitHigh;                      // 内环上饱和（当拍量）
_bSatLow := fbInner.bLimitLow;                        // 内环下饱和（当拍量）
rtReset(CLK := bReset);                               // 复位沿（每拍必调）
tonSatHiTo(IN := bEnable AND _bSatHigh, PT := tSatTo);    // 上饱和确认（每拍必调）
tonSatLoTo(IN := bEnable AND _bSatLow, PT := tSatTo);     // 下饱和确认（每拍必调）

(* —— 段 1：单拍量预清零（锁存量 _uFault/_bHiLat/_bLoLat/_bCfgBad 不入清单，禁同拍抹除） —— *)
_uInfo := 16#0000_0000;             // 信息码每拍重算
bFreeze := FALSE;                   // 冻结出口缺省 FALSE
bMirror := FALSE;                   // 镜像出口缺省 FALSE
nErrId := 16#0000_0000;             // 事件码缺省无事件

(* —— 段 2：复位沿 + 组态域闸（当拍量判据） —— *)
IF rtReset.Q THEN                   // rtReset.Q = 当拍量
    _bHiLat := FALSE;               // 清上饱和锁存位
    _bLoLat := FALSE;               // 清下饱和锁存位
    _bCfgBad := FALSE;              // 清组态锁存位
    _uFault := 16#0000_0000;        // 清故障锁存码
END_IF
IF fInnerMax <= fInnerMin THEN
    _uFault := 16#0002_03AB;        // 故障级：组态非法（限幅颠倒）
    _bCfgBad := TRUE;
END_IF

(* —— 段 3：限幅镜像（仅组态有效且使能相生效；R242：仅外环 bTrack=FALSE 相写入） —— *)
IF bEnable AND (NOT _bCfgBad) AND (NOT fbOuter.bTrack) THEN
    fbOuter.rOutMin := fInnerMin;   // 外环下限镜像内环
    fbOuter.rOutMax := fInnerMax;   // 外环上限镜像内环
    bMirror := TRUE;                // 镜像生效标志
    IF NOT _bMirrorSent THEN
        _uInfo := 16#0002_0491;     // 信息级：镜像钳制生效沿
        _bMirrorSent := TRUE;       // 沿单发
    END_IF
END_IF

(* —— 段 4：饱和锁存与解除（判据当拍量；解除式全当拍量，R240 落地） —— *)
IF tonSatHiTo.Q AND (NOT _bHiLat) THEN
    _uFault := 16#0002_03AC;        // 故障级：上饱和持续锁存
    _bHiLat := TRUE;
END_IF
IF tonSatLoTo.Q AND (NOT _bLoLat) THEN
    _uFault := 16#0002_03AD;        // 故障级：下饱和持续锁存
    _bLoLat := TRUE;
END_IF
(* 解除式逐 BOOL 标注（R240）：rtReset.Q = 当拍量；_bSatHigh/_bSatLow = 当拍量；
   均不含锁存量（_bHiLat/_bLoLat），解除边真实可达。 *)
IF rtReset.Q AND (NOT _bSatHigh) AND (NOT _bSatLow) AND (NOT _bCfgBad) THEN
    _bHiLat := FALSE;               // 清上饱和锁存位（锁存量，仅此当拍量解除沿可清）
    _bLoLat := FALSE;               // 清下饱和锁存位（锁存量，仅解除沿可清）
    _uFault := 16#0000_0000;        // 清故障锁存码（锁存量，仅本当拍量解除沿可清）
END_IF

(* —— 段 5：外环输出非有限防御兜底（NaN 自反判） —— *)
IF (fbOuter.fOut <> fbOuter.fOut) OR ((fbOuter.fOut - fbOuter.fOut) <> (fbOuter.fOut - fbOuter.fOut)) THEN
    _uFault := 16#0002_03AE;        // 故障级：外环输出非有限
    _bHiLat := TRUE;                // 并入聚合锁存（安全侧）
END_IF

(* —— 段 6：外环积分冻结联动（R242：bExtTrack 相冻结让位；冻结经跟踪机制承载） —— *)
IF bEnable AND (NOT _bCfgBad) AND (_bSatHigh OR _bSatLow) AND (NOT bExtTrack) THEN
    fbOuter.bTrack := TRUE;         // 冻结：跟踪机制接管
    fbOuter.fTrackValue := fbOuter.fOut;    // 跟踪值 = 当前输出（保持不积分）
    bFreeze := TRUE;                // 冻结生效标志
    IF NOT _bFreezePrev THEN
        _uInfo := 16#0002_0492;     // 信息级：冻结激活沿
    END_IF
ELSIF bEnable AND (NOT _bCfgBad) AND bExtTrack THEN
    fbOuter.bTrack := TRUE;         // 外部跟踪直通（调用方所有权）
    fbOuter.fTrackValue := fExtTrackVal;    // 外部跟踪值
    IF (_bSatHigh OR _bSatLow) THEN
        _uInfo := 16#0002_0494;     // 信息级：冻结请求被外部跟踪让位
    END_IF
ELSE
    fbOuter.bTrack := FALSE;        // 解除跟踪（恢复 PID 自主积分）
    IF _bFreezePrev THEN
        _uInfo := 16#0002_0493;     // 信息级：冻结解除恢复沿
    END_IF
END_IF

(* —— 段 7：出口单点映射（锁存码回放，禁同拍抹除） —— *)
IF (_bHiLat OR _bLoLat OR _bCfgBad) THEN
    nErrId := _uFault;              // 故障锁存码回放
    bFreeze := FALSE;               // 故障期冻结出口强制 FALSE（安全侧）
    bMirror := FALSE;               // 故障期镜像出口强制 FALSE（安全侧）
    fbOuter.bTrack := FALSE;        // 故障期跟踪标志与钳制同步释放（v1.0.1 名实一致，R191）
ELSE
    nErrId := _uInfo;               // 信息码
END_IF
bError := _bHiLat OR _bLoLat OR _bCfgBad;   // 故障标志与锁存位同源
_bFreezePrev := bFreeze;            // 冻结解除沿判据快照

END_FUNCTION_BLOCK

(* ---- FB_DL_ChwDifferentialPressure.st ---- *)
// =====================================================================
// FB_DL_ChwDifferentialPressure.st
// 冷冻水差压旁通控制（压差平滑 + 设定值重置限速 + PID 指令注入 + 阀位限幅）
// CHW differential pressure bypass control with smoothing and valve clamp
// 所属子库: DL_Algo    版本: v1.0.0    兼容: CODESYS V3.5+ / TwinCAT 3 / 汇川 InoProShop
// 码位: 16#0002_372E ~ 16#0002_3732 (本件独占 5 槽, 勿复用)
// 溯源: 道莅 clean-room 防御性实现
//       来源组标签: hvac, chw, differential-pressure, pid
// 修改记录: R30 初版 (ROUND_PLAN_R30 序 18)
// 分层声明: 压差平滑组合消费 DL_MathData 的 FB_DL_MovingAverage 实例;
//           设定值重置限速组合消费 DL_Algo 的 FB_DL_RateLimiter 实例
//           （斜坡防水锤）; PID 闭环本身不内联, 控制件阀位指令输出经引脚注入
// =====================================================================
FUNCTION_BLOCK FB_DL_ChwDifferentialPressure
VAR_INPUT
    bEnable        : BOOL  := FALSE;   // 使能 / Enable
    fDp_kPa        : REAL  := 0.0;     // 供回水压差 0~400 kPa / Supply-return dP [kPa]
    fDpSet_kPa     : REAL  := 120.0;   // 压差设定值 0~400 kPa / dP setpoint [kPa]
    fPidOut_Pct    : REAL  := 0.0;     // PID 阀位指令注入（控制件 fOut 语义）/ PID valve command injected [pct]
    fValveMin_Pct  : REAL  := 0.0;     // 阀位下限 0~100 百分比 / Valve lower limit [pct]
    fValveMax_Pct  : REAL  := 100.0;   // 阀位上限 0~100 百分比 / Valve upper limit [pct]
    fResetRate_kPa_s: REAL := 5.0;     // 设定值重置限速 0~100 kPa/s, 0 = 不限 / Setpoint reset rate [kPa/s]
END_VAR
VAR_OUTPUT
    fValveOut_Pct  : REAL  := 0.0;    // 旁通阀位输出 / Bypass valve output [pct]
    fDpSmooth_kPa  : REAL  := 0.0;    // 平滑后压差 / Smoothed dP [kPa]
    bByPassActive  : BOOL  := FALSE;  // 旁通投入标志 / Bypass active flag
    eErr           : UDINT := 16#0002_372E;  // 错误码 / Error code
END_VAR
VAR
    movAvg      : FB_DL_MovingAverage;  // 压差平滑实例（组合消费）/ Smoothing instance, composed
    ratSet      : FB_DL_RateLimiter;    // 设定值限速实例（组合消费）/ Setpoint rate limiter instance
    bCfgErr     : BOOL  := FALSE;   // 组态非法标记 / Configuration error flag
    bInFErr     : BOOL  := FALSE;   // 输入非有限标记 / Input non-finite flag
    bSatInfo    : BOOL  := FALSE;   // 阀位限幅饱和信息标记 / Valve saturation info flag
    fValveHold  : REAL  := 0.0;     // 阀位保持量（非有限拍保持）/ Valve hold value [pct]
    fValveCmd   : REAL  := 0.0;     // 阀位指令临时量 / Valve command temporary [pct]
    fSetUse     : REAL  := 0.0;     // 限速后设定值（诊断保持）/ Rate-limited setpoint [kPa]
END_VAR

// ---------------------------------------------------------------------
// 代码位表（本件独占, 勿复用）:
//   16#0002_372E 信息 旁通控制正常
//   16#0002_372F 故障 输入非有限（压差或 PID 指令注入非有限, 阀位保持上拍值,
//                不新增动作）; 解除式 = 输入恢复有限
//   16#0002_3730 故障 组态非法（设定值越出 0~400 kPa, 阀限幅越域或倒置,
//                重置速率越出 0~100 kPa/s）; 解除式 = 恢复合法组态
//   16#0002_3731 信息 阀位限幅饱和（PID 指令越出阀限幅, 已钳位输出）
//   16#0002_3732 信息 待机未使能（阀位回下限, 旁通关闭安全侧）
// ---------------------------------------------------------------------

// ---- 组态闸 / Configuration gate ----
bCfgErr := FALSE;
IF (fDpSet_kPa <> fDpSet_kPa) OR (fDpSet_kPa < 0.0) OR (fDpSet_kPa > 400.0) THEN
    bCfgErr := TRUE;                // 设定值越域 / Setpoint out of domain
END_IF
IF (fValveMin_Pct <> fValveMin_Pct) OR (fValveMin_Pct < 0.0) OR (fValveMin_Pct > 100.0) THEN
    bCfgErr := TRUE;                // 下限越域 / Lower limit out of domain
END_IF
IF (fValveMax_Pct <> fValveMax_Pct) OR (fValveMax_Pct < 0.0) OR (fValveMax_Pct > 100.0) THEN
    bCfgErr := TRUE;                // 上限越域 / Upper limit out of domain
END_IF
IF (NOT bCfgErr) AND (fValveMin_Pct >= fValveMax_Pct) THEN
    bCfgErr := TRUE;                // 阀限幅倒置 / Inverted valve limits
END_IF
IF (fResetRate_kPa_s <> fResetRate_kPa_s) OR (fResetRate_kPa_s < 0.0) OR (fResetRate_kPa_s > 100.0) THEN
    bCfgErr := TRUE;                // 重置速率越域 / Reset rate out of domain
END_IF

// ---- 输入非有限判 / Input finite judge ----
bInFErr := (fDp_kPa <> fDp_kPa) OR (ABS(fDp_kPa) >= 1.0E12)
        OR (fPidOut_Pct <> fPidOut_Pct) OR (ABS(fPidOut_Pct) >= 1.0E12);

// ---- 压差平滑消费（组合实例调用）/ Smoothing via composed instance ----
movAvg(fInput := fDp_kPa, nWindowSize := 8,
       bSample := bEnable AND (NOT bInFErr) AND (NOT bCfgErr),
       bEnable := bEnable, bReset := FALSE);
fDpSmooth_kPa := movAvg.fAverage;   // 平滑压差输出 / Smoothed dP output

// ---- 设定值重置限速消费（组合实例调用, 斜坡防水锤）/ Setpoint rate limit ----
ratSet(bEnable := bEnable AND (NOT bCfgErr), fIn := fDpSet_kPa,
       fRateUp := fResetRate_kPa_s, fRateDown := fResetRate_kPa_s,
       bTrack := (NOT bEnable), fTrackValue := fDpSet_kPa,
       tSampleTime := T#100MS);
fSetUse := ratSet.fOut;             // 限速后设定值保持（供上位诊断）/ Held setpoint for diagnostics

// ---- 待机安全侧: 阀位回下限（旁通关闭）/ Standby: valve to lower limit ----
IF NOT bEnable THEN
    fValveOut_Pct := fValveMin_Pct; // 关闭旁通 / Close bypass
    fValveHold := fValveMin_Pct;    // 保持量同步 / Sync hold
    bByPassActive := FALSE;         // 旁通退出 / Bypass off
    eErr := 16#0002_3732;           // 待机码 / Standby code
ELSIF bInFErr OR bCfgErr THEN
    // 非有限或组态非法: 阀位保持上拍值, 不新增动作 / Hold valve, no new action
    fValveOut_Pct := fValveHold;
    bByPassActive := FALSE;
    IF bCfgErr THEN
        eErr := 16#0002_3730;       // 组态码 / Config code
    ELSE
        eErr := 16#0002_372F;       // 非有限码 / Non-finite code
    END_IF
ELSE
    // ---- 阀位指令限幅输出 / Valve command with clamping ----
    fValveCmd := fPidOut_Pct;       // PID 指令注入 / Injected PID command
    bSatInfo := FALSE;
    IF fValveCmd > fValveMax_Pct THEN
        fValveCmd := fValveMax_Pct; // 上限钳位 / Clamp upper
        bSatInfo := TRUE;           // 置饱和信息 / Set saturation info
    END_IF
    IF fValveCmd < fValveMin_Pct THEN
        fValveCmd := fValveMin_Pct; // 下限钳位 / Clamp lower
        bSatInfo := TRUE;
    END_IF
    fValveOut_Pct := fValveCmd;     // 阀位输出 / Valve output
    fValveHold := fValveCmd;        // 更新保持量 / Update hold
    // 旁通投入判（容差比较, 浮点禁直接判等）/ Bypass active with margin
    bByPassActive := (fValveOut_Pct - fValveMin_Pct) > 0.1;
    IF bSatInfo THEN
        eErr := 16#0002_3731;       // 饱和信息 / Saturation info
    ELSE
        eErr := 16#0002_372E;       // 正常 / Normal
    END_IF
END_IF

END_FUNCTION_BLOCK

(* ---- FB_DL_ChwDifferentialPressureReset.st ---- *)
(*
  FB_DL_ChwDifferentialPressureReset  —  冷冻水压差重置（阀位反馈反算设定 + 死区保持） / Chilled-water differential-pressure reset by valve-position back-calculation with deadband hold
  分类 Category : DL_Algo
  版本 Version  : 1.0.0
  来源 Source   : t1-2-oscat-building — 楼宇冷冻水压差重置算法族深化
  溯源 Origin   : 道莅 clean-room 实现；阀位反馈线性反算压差设定 + 死区保持 + 限速为公开水系统节能算法，未复制任何源码行
  功能 Function : 1) 反算：fDpSpRawKpa = fDpBaseKpa + fDpGainKpaPerPct × (fValveFbPct - fValveTargetPct)
                  （阀位大于目标阀位意味着压差不足 → 抬高设定）；
                  2) 死区保持：|反算值 - 当前输出| < fDeadbandKpa 时输出保持不变；
                  3) 限速：单次调用变化量不超过 fMaxStepKpa（与逐周期积分爬坡不同，本件为
                  反算直给的限速钳制，超限时按步长逼近）；
                  4) 硬限幅 [fDpMinKpa, fDpMaxKpa]，限幅后二次复核；
                  5) 本件只有故障码、无信息码（派单硬约束）。
  接口 Interface: 输入阀位反馈/目标阀位/基准/增益/死区/步长/上下限；输出压差设定
  边界 Boundary : ① 组态闸：fDpMaxKpa <= fDpMinKpa、fMaxStepKpa <= 0.0、fDeadbandKpa < 0.0、
                  fDpGainKpaPerPct <= 0.0 → 0388 锁存；
                  ② 阀位与压差量非有限（NaN 自反 + Inf 差值自减）→ 0388 锁存，设定冻结保持
                  （R191：语义为冻结保持，非降级置标志）；
                  ③ 浮点判据全容差式；④ 仅一个 R_TRIG 复位沿，段 0 无条件调用；
                  ⑤ 故障相迁出唯一路径 = bReset 上升沿；⑥ 零全局耦合（无 GVL / %I %Q %M）。
  依赖 Depends  : Standard.library（R_TRIG）
  码表 Error codes（Algo 段 0002，故障窗口 0388；本件无信息码）:
    16#0002_0388 故障级：压差重置故障总码（组态非法 / 阀位或压差量非有限），
                 锁存至 bReset 上升沿；归因见 eCause，不新增码位（派单硬约束单码）
  修订历史 Revision :
    2026-11-19  v1.0.0  R43 首版（批次 3 · 序号 12）
*)

TYPE E_DL_CdpState :
(
    eIdle   := 0,     // 未使能：设定冻结 / Idle, setpoint frozen
    eRun    := 10,    // 反算运行中 / Back-calculation active
    eFault  := 90     // 故障锁存相（设定冻结保持） / Fault latched, setpoint frozen
);
END_TYPE

TYPE E_DL_CdpCause :
(
    eNone       := 0, // 无故障成因 / No cause
    eCfgIllegal := 1, // 组态非法 / Illegal configuration
    eNonFinite  := 2  // 输入非有限 / Non-finite input
);
END_TYPE

FUNCTION_BLOCK FB_DL_ChwDifferentialPressureReset
VAR_INPUT
    fValveFbPct       : REAL := 0.0;     // 末端阀位反馈 [%]，0~100 / Terminal valve feedback
    fValveTargetPct   : REAL := 85.0;    // 目标阀位 [%]，开区间 (0,100) / Target valve position
    fDpBaseKpa        : REAL := 150.0;   // 压差基准 [kPa] / Base differential pressure
    fDpGainKpaPerPct  : REAL := 2.0;     // 反算增益 [kPa/%]，域 > 0 / Back-calculation gain
    fDeadbandKpa      : REAL := 3.0;     // 死区 [kPa]，域 >= 0 / Deadband
    fMaxStepKpa       : REAL := 10.0;    // 单次限速步长 [kPa]，域 > 0 / Rate limit step
    fDpMinKpa         : REAL := 50.0;    // 压差设定下限 [kPa] / Setpoint low limit
    fDpMaxKpa         : REAL := 300.0;   // 压差设定上限 [kPa] / Setpoint high limit
    fDpInitKpa        : REAL := 150.0;   // 设定初值（使能沿装载） [kPa] / Initial setpoint
    bEnable           : BOOL := FALSE;   // 反算使能（电平）[-] / Reset enable
    bReset            : BOOL := FALSE;   // 复位命令，上升沿清故障 [-] / Reset edge
END_VAR
VAR_OUTPUT
    eState            : E_DL_CdpState;   // 状态出口，段 6 单点映射 / State outlet
    eCause            : E_DL_CdpCause;   // 故障成因出口（R190） / Fault cause outlet
    fDpSpKpa          : REAL;            // 压差设定输出 [kPa] / Differential pressure setpoint
    fDpSpRawKpa       : REAL;            // 反算原始值镜像 [kPa] / Raw back-calculated value
    bDbHold           : BOOL;            // 死区保持镜像 [-] / Deadband hold mirror
    bError            : BOOL;            // 故障锁存标志 [-] / Fault latch flag
    nErrId            : UDINT;           // 故障码，0 = 无故障（本件无信息码） / Fault code only
END_VAR
VAR
    _eState           : E_DL_CdpState := E_DL_CdpState.eIdle;   // 内部相位（CASE 唯一写入目标） / Internal phase
    _eCause           : E_DL_CdpCause := E_DL_CdpCause.eNone;   // 故障成因锁存（锁存量） / Latched cause
    rtEnable          : R_TRIG;          // 使能沿实例，每周期无条件调用 / Enable edge
    rtReset           : R_TRIG;          // 复位沿实例，每周期无条件调用 / Reset edge
    _fSp              : REAL;            // 设定保持槽（持久） / Setpoint holding slot
    _fRawKpa          : REAL;            // 反算原始值 [kPa]（当拍量） / Raw value
    _fCandKpa         : REAL;            // 限幅-限速后候选 [kPa]（当拍量） / Candidate value
    _bDbHoldOn        : BOOL;            // 死区保持当拍量 [-] / Deadband hold flag
    _bNonFin          : BOOL;            // 输入非有限当拍量 [-] / Non-finite input
    _bCfgBad          : BOOL;            // 组态非法当拍量 [-] / Config illegal
    _bFault           : BOOL;            // 故障锁存位（锁存量） / Latched fault bit
    _uFault           : UDINT;           // 故障码锁存（锁存量） / Latched fault code
END_VAR

(* —— 段 0：沿实例无条件周期刷新 + 当拍量判据 —— *)
_fRawKpa := fDpBaseKpa + fDpGainKpaPerPct * (fValveFbPct - fValveTargetPct);   // 阀位反算压差 [kPa] / Back-calculated pressure
_bNonFin := (fValveFbPct <> fValveFbPct) OR (fDpBaseKpa <> fDpBaseKpa)
         OR ((fValveFbPct - fValveFbPct) <> (fValveFbPct - fValveFbPct))
         OR ((fDpBaseKpa - fDpBaseKpa) <> (fDpBaseKpa - fDpBaseKpa));           // NaN 自反 + Inf 差值自减 / NaN and Inf
_bCfgBad := (fDpMaxKpa <= fDpMinKpa) OR (fMaxStepKpa <= 0.0) OR (fDeadbandKpa < 0.0)
            OR (fDpGainKpaPerPct <= 0.0) OR (fValveTargetPct <= 0.0) OR (fValveTargetPct >= 100.0);   // 组态非法当拍量 / Config illegal
rtEnable(CLK := bEnable);                                                       // 使能沿，每拍必调 / Enable edge
rtReset(CLK := bReset);                                                         // 复位沿，每拍必调 / Reset edge

(* —— 段 1：单拍量预清零（锁存量与设定保持槽不入清单） —— *)
fDpSpRawKpa := 0.0;                // 反算镜像缺省 0 / Raw mirror default
bDbHold := FALSE;                  // 死区镜像缺省 FALSE / Deadband default
nErrId := 16#0000_0000;            // 故障码缺省无故障 / Fault code default

(* —— 段 2：复位沿 + 组态域闸 —— *)
IF rtReset.Q THEN                              // rtReset.Q = 当拍量 / current scan
    _bFault := FALSE;                          // 清故障锁存位（锁存量） / Clear fault latch
    _uFault := 16#0000_0000;                   // 清故障锁存码（锁存量） / Clear fault code
    _eCause := E_DL_CdpCause.eNone;            // 清成因（锁存量） / Clear cause
    IF _eState = E_DL_CdpState.eFault THEN
        _eState := E_DL_CdpState.eIdle;        // 故障相迁出：回未使能 / Fault exit to idle
    END_IF
END_IF
IF _bCfgBad THEN                               // 组态域闸 / Config gate
    _uFault := 16#0002_0388;                   // 故障级：重置故障总码 / Algo fault code
    _eCause := E_DL_CdpCause.eCfgIllegal;      // 归因：组态非法 / Cause: illegal config
    _bFault := TRUE;                           // 标志与码位配对（R45） / Flag paired with code
END_IF
IF (NOT _bFault) AND _bNonFin THEN             // 非有限锁存 / Non-finite latch
    _uFault := 16#0002_0388;
    _eCause := E_DL_CdpCause.eNonFinite;       // 归因：非有限 / Cause: non-finite
    _bFault := TRUE;
END_IF

(* —— 段 3：反算 + 死区 + 限速 + 限幅（仅运行相且无故障） —— *)
IF (NOT _bFault) AND (_eState = E_DL_CdpState.eRun) THEN
    _fCandKpa := _fRawKpa;                                 // 候选 = 反算原始值 / Candidate from raw
    IF _fCandKpa < fDpMinKpa THEN                          // 下限钳制 / Low clamp
        _fCandKpa := fDpMinKpa;
    ELSIF _fCandKpa > fDpMaxKpa THEN                       // 上限钳制 / High clamp
        _fCandKpa := fDpMaxKpa;
    END_IF
    IF ABS(_fCandKpa - _fSp) < fDeadbandKpa THEN           // 死区内保持（容差式） / Deadband hold
        _bDbHoldOn := TRUE;
    ELSIF (_fCandKpa - _fSp) > fMaxStepKpa THEN            // 向上限速 / Upward rate limit
        _fSp := _fSp + fMaxStepKpa;
    ELSIF (_fSp - _fCandKpa) > fMaxStepKpa THEN            // 向下限速 / Downward rate limit
        _fSp := _fSp - fMaxStepKpa;
    ELSE
        _fSp := _fCandKpa;                                 // 直接跟随反算值 / Follow candidate
    END_IF
    IF _fSp < fDpMinKpa THEN                               // 限速后二次下限复核 / Post-limit low check
        _fSp := fDpMinKpa;
    ELSIF _fSp > fDpMaxKpa THEN                            // 限速后二次上限复核 / Post-limit high check
        _fSp := fDpMaxKpa;
    END_IF
END_IF

(* —— 段 4：故障解除式（R240；全当拍量）：rtReset.Q / NOT _bCfgBad / NOT _bNonFin —— *)
IF rtReset.Q AND (NOT _bCfgBad) AND (NOT _bNonFin) THEN
    _bFault := FALSE;                          // 清故障锁存位（锁存量） / Clear fault latch
    _uFault := 16#0000_0000;                   // 清故障锁存码（锁存量） / Clear fault code
    _eCause := E_DL_CdpCause.eNone;            // 清成因（锁存量） / Clear cause
END_IF

(* —— 段 4A：故障锁存相位迁移闸（设定冻结保持） —— *)
IF _bFault AND (_eState <> E_DL_CdpState.eFault) THEN
    _eState := E_DL_CdpState.eFault;           // 锁存即入故障相 / Latch enters fault phase
END_IF

(* —— 段 5：相位机（CASE 全覆盖 + ELSE 兜底） —— *)
CASE _eState OF

E_DL_CdpState.eIdle:
    IF rtEnable.Q AND (NOT _bFault) THEN       // 使能上升沿：装载初值并钳制 / Enable edge loads initial value
        _fSp := fDpInitKpa;                    // 装载初值 / Load initial setpoint
        IF _fSp < fDpMinKpa THEN               // 初值下限钳制 / Initial low clamp
            _fSp := fDpMinKpa;
        ELSIF _fSp > fDpMaxKpa THEN            // 初值上限钳制 / Initial high clamp
            _fSp := fDpMaxKpa;
        END_IF
        _eState := E_DL_CdpState.eRun;         // 进运行相 / Enter run
    END_IF

E_DL_CdpState.eRun:
    IF NOT bEnable THEN                        // 撤使能：设定冻结，回未使能 / Disable: freeze and idle
        _eState := E_DL_CdpState.eIdle;
    END_IF

E_DL_CdpState.eFault:
    ;                                          // 故障相：设定冻结保持，仅段 4 复位沿可迁出 / Frozen, reset only

ELSE
    _uFault := 16#0002_0388;                   // 故障级：非法相位兜底（归并总码） / Illegal phase fallback
    _eCause := E_DL_CdpCause.eCfgIllegal;      // 归因：相位非法归并组态 / Cause: phase illegal
    _bFault := TRUE;
    _eState := E_DL_CdpState.eFault;           // 强制回故障相 / Force fault phase

END_CASE

(* —— 段 6：出口单点映射（名实同源；锁存码回放） —— *)
fDpSpKpa := _fSp;                              // 设定值出口 / Setpoint outlet
IF _bFault THEN
    nErrId := _uFault;                         // 故障锁存码回放 / Replay latched code
    fDpSpRawKpa := 0.0;                        // 故障相反算镜像强制 0 / Raw mirror forced zero
    bDbHold := FALSE;                          // 故障相死区镜像强制 FALSE / Deadband forced false
ELSE
    nErrId := 16#0000_0000;                    // 无故障：本件无信息码 / No fault, no info code
    fDpSpRawKpa := _fRawKpa;                   // 反算镜像 / Raw mirror
    bDbHold := _bDbHoldOn;                     // 死区镜像 / Deadband mirror
END_IF
bError := _bFault;                             // 故障标志同源 / Flag from latch
eState := _eState;                             // 状态出口 / State outlet
eCause := _eCause;                             // 成因出口 / Cause outlet

END_FUNCTION_BLOCK

(* ---- FB_DL_CoatingThicknessCtrl.st ---- *)
// =====================================================================
// FB_DL_CoatingThicknessCtrl.st
// 涂布面密度闭环控制（一阶滤波 + 纯滞后补偿 + 积分型无差调节）
// Coating weight closed-loop control FB
// 码位: 16#0002_371A ~ 16#0002_371E (本件独占 5 槽)
// 修改记录: R29 初版 (按 DISPATCH_R29 序 4)
// =====================================================================
FUNCTION_BLOCK FB_DL_CoatingThicknessCtrl
VAR_INPUT
    bEnable            : BOOL  := FALSE;   // 使能，FALSE 冻结输出 / Enable, freeze outputs when FALSE
    bStart             : BOOL  := FALSE;   // 上升沿投入闭环 / Start on rising edge
    bReset             : BOOL  := FALSE;   // 复位故障，仅 eFault 生效 / Fault reset
    bMeasValid         : BOOL  := FALSE;   // 测厚数据有效 / Measurement valid
    fMeas_gsm          : REAL  := 0.0;     // 实测面密度 0~500 g/m² / Measured coat weight [g/m2]
    fSp_gsm            : REAL  := 120.0;   // 面密度设定 1~500 g/m² / Setpoint [g/m2]
    fBandPct           : REAL  := 0.5;     // 死区带 0~5 % / Dead band [%]
    fGain_mm_per_gsm   : REAL  := 0.01;    // 间隙-面密度增益 0.0001~1 mm/(g/m²) / Gap gain [mm/(g/m2)]
    fGapInit_mm        : REAL  := 0.250;   // 初始间隙 0.05~2.0 mm / Initial gap [mm]
    fTrimMax_mm        : REAL  := 0.100;   // 相对初始间隙最大修正 0.001~1.0 mm / Max trim [mm]
    fRateMax_mm_s      : REAL  := 0.005;   // 修正速率上限 >0 mm/s / Trim rate limit [mm/s]
    tDeadTime          : TIME  := T#30S;   // 纯滞后 T#1S~T#300S / Dead time [s]
    tCycle             : TIME  := T#100MS; // 采样周期 T#10MS~T#5S / Sample cycle [s]
END_VAR
VAR_OUTPUT
    fGapCmd_mm         : REAL;             // 模头间隙命令 0.05~2.0 mm / Gap command [mm]
    fDev_gsm           : REAL;             // 滞后补偿后偏差 g/m² / Delayed deviation [g/m2]
    fTrim_mm           : REAL;             // 当前累计修正 mm / Accumulated trim [mm]
    bInBand            : BOOL;             // 偏差在带内 / Within dead band
    bActive            : BOOL;             // 闭环投入中 / Loop active
    eState             : E_DL_CoatingState; // 状态 / State
    eErr               : UDINT;            // 错误码 / Error code
END_VAR
VAR
    rtrigStart         : R_TRIG;           // 启动上升沿检测 / Start rising-edge detector
    fFilt_gsm          : REAL;             // 一阶滤波后测厚值 / Filtered measurement [g/m2]
    fDevNow_gsm        : REAL;             // 本拍新鲜偏差 / Fresh deviation this cycle [g/m2]
    aDelayQ            : ARRAY[0..2999] OF REAL; // 延时队列（偏差历史）/ Delay queue of deviations [g/m2]
    uQHead             : UDINT;            // 队列写指针 / Queue write pointer
    uQLen              : UDINT;            // 队列有效长度 / Queue valid length
    uQLenCfg           : UDINT;            // 组态队列长度（CEIL 后）/ Configured queue length
    uIdx               : UDINT;            // 循环下标 / Loop index
    fRateStep          : REAL;             // 单拍速率步长 / Rate step per cycle [mm]
    fTrimNew           : REAL;             // 修正后临时累计值 / Tentative new trim [mm]
    fBandAbs           : REAL;             // 死区绝对带宽 / Absolute dead band [g/m2]
    tCycleS            : REAL;             // 周期秒值（钳 ≥0.01）/ Cycle in seconds, clamped [s]
    tDeadS             : REAL;             // 滞后秒值 / Dead time in seconds [s]
    xFirstScan         : BOOL := TRUE;     // 首扫标记 / First-scan flag
    tCyclePrev         : TIME  := T#0MS;   // 上拍周期快照 / Previous cycle snapshot
END_VAR

// ---------------------------------------------------------------------
// 代码位表（本件独占，勿复用）:
//   16#0002_371A 信息 闭环运行正常 / 带内不动作
//   16#0002_371B 故障 输入非有限，或 tDeadTime/tCycle 非法（0 或超出域）
//   16#0002_371C 故障 fGain/fTrimMax/fRateMax/fSp 组态错（≤0）
//   16#0002_371D 信息 修正触限 → 停止同向积分，eState=eLimit
//   16#0002_371E 信息 测厚无效 → 冻结积分、输出保持、bActive=FALSE
// ---------------------------------------------------------------------

// ---- 时间参数转秒（TIME/1000 毫秒基准）/ Convert times to seconds ----
tCycleS := TIME_TO_REAL(tCycle) / 1000.0;   // 周期秒值 / Cycle seconds [s]
tDeadS  := TIME_TO_REAL(tDeadTime) / 1000.0; // 滞后秒值 / Dead-time seconds [s]
IF tCycleS < 0.01 THEN
    tCycleS := 0.01;    // 钳下限防步长爆炸 / Clamp minimum 10 ms
END_IF

// ---- 组态合法性检查（故障级，锁存于 eFault）/ Configuration validity check ----
IF (tCycle = T#0MS) OR (tDeadTime = T#0MS)
   OR (tDeadS > 300.0) OR (tDeadS < 1.0)
   OR (tCycleS > 5.0)
   OR (fMeas_gsm <> fMeas_gsm) OR (ABS(fMeas_gsm) >= 1.0E12)
   OR (fSp_gsm <> fSp_gsm) OR (ABS(fSp_gsm) >= 1.0E12) THEN
    // 非有限或时域非法 / Non-finite or invalid time domain
    IF eState <> E_DL_CoatingState.eFault THEN
        eState := E_DL_CoatingState.eFault;  // 进入故障态（锁存）/ Enter latched fault
    END_IF
    bActive  := FALSE;          // 闭环退出 / Loop inactive
    eErr     := 16#0002_371B;   // 故障码 / Fault code
    // 故障态输出保持，不推进 / Hold outputs, no advance
    RETURN;                     // 本拍结束 / End of cycle
END_IF

// ---- 组态错闸（故障级）/ Configuration fault gate ----
IF (fGain_mm_per_gsm <= 0.0) OR (fTrimMax_mm <= 0.0)
   OR (fRateMax_mm_s <= 0.0) OR (fSp_gsm <= 0.0) THEN
    IF eState <> E_DL_CoatingState.eFault THEN
        eState := E_DL_CoatingState.eFault;  // 进入故障态（锁存）/ Enter latched fault
    END_IF
    bActive := FALSE;           // 闭环退出 / Loop inactive
    eErr    := 16#0002_371C;    // 故障码 / Fault code
    RETURN;                     // 本拍结束 / End of cycle
END_IF

// ---- 延时队列长度组态 = CEIL(tDeadTime/tCycle)，上限 3000 拍 / Delay queue length config ----
uQLenCfg := REAL_TO_UDINT(CEIL(tDeadS / tCycleS));  // 拍数 / Queue length in cycles
IF uQLenCfg > 3000 THEN
    uQLenCfg := 3000;           // 超限按 3000 防内存爆 / Cap at 3000
    IF eState <> E_DL_CoatingState.eFault THEN
        eState := E_DL_CoatingState.eFault;  // 故障锁存 / Latch fault
    END_IF
    bActive := FALSE;           // 闭环退出 / Loop inactive
    eErr    := 16#0002_371B;    // 故障码 / Fault code
    RETURN;                     // 本拍结束 / End of cycle
END_IF
IF uQLenCfg = 0 THEN
    uQLenCfg := 1;              // 至少 1 拍防零长度 / Minimum 1 cycle
END_IF

// ---- 故障复位（仅 eFault 生效）/ Fault reset only in fault state ----
IF (eState = E_DL_CoatingState.eFault) AND bReset THEN
    eState := E_DL_CoatingState.eIdle;  // 回空闲态 / Back to idle
    fTrim_mm := 0.0;            // 清累计修正 / Clear trim
    uQLen := 0;                 // 清延时队列 / Clear delay queue
    uQHead := 0;                // 指针归零 / Reset pointer
END_IF

// ---- 首扫初始化（R16 首扫纪律）/ First-scan initialization ----
IF xFirstScan THEN
    fGapCmd_mm := fGapInit_mm;  // 首扫置初始间隙 / Init gap on first scan
    fFilt_gsm  := fSp_gsm;      // 滤波器初值取设定 / Filter init at setpoint
    xFirstScan := FALSE;        // 清首扫标记 / Clear flag
    tCyclePrev := tCycle;       // 记录周期 / Record cycle
END_IF

// ---- 周期变化检测：清队列并重填当前偏差 / Cycle change: flush queue and refill ----
IF (tCyclePrev <> tCycle) AND (NOT xFirstScan) THEN
    FOR uIdx := 0 TO 2999 DO
        aDelayQ[uIdx] := 0.0;   // 清空历史脏值 / Clear stale history
    END_FOR
    fFilt_gsm := fSp_gsm;       // 滤波器重新对齐设定 / Re-align filter
    uQLen := 0;                 // 清队列长度 / Reset length
    uQHead := 0;                // 指针归零 / Reset pointer
    tCyclePrev := tCycle;       // 更新周期快照 / Update snapshot
END_IF

// ---- 启动沿：仅 eIdle 可进 eRun，非沿不重复初始化 / Start edge: idle to run only ----
rtrigStart(CLK := bStart);      // 沿检测无条件周期刷新 / Unconditional per-cycle refresh
IF rtrigStart.Q AND (eState = E_DL_CoatingState.eIdle) AND bEnable THEN
    eState    := E_DL_CoatingState.eRun;  // 投入闭环 / Activate loop
    fTrim_mm  := 0.0;           // 清累计修正 / Clear trim
    fGapCmd_mm := fGapInit_mm;  // 间隙回初始值 / Reset gap to initial
    fFilt_gsm := fSp_gsm;       // 滤波器重新对齐 / Re-align filter
    uQLen := 0;                 // 清延时队列 / Clear queue
    uQHead := 0;                // 指针归零 / Reset pointer
END_IF

// ---- 输出默认量 / Default per-cycle outputs ----
bActive := FALSE;               // 默认非投入 / Default inactive
bInBand := FALSE;               // 默认带外 / Default out of band

// ---- 状态机 / State machine ----
CASE eState OF

    E_DL_CoatingState.eIdle:    // 空闲态 / Idle state
        fGapCmd_mm := fGapInit_mm;  // 间隙保持初始 / Hold initial gap
        fTrim_mm   := 0.0;          // 修正清零 / Trim zero
        eErr       := 16#0002_371A; // 信息级：正常空闲 / Info: idle normal

    E_DL_CoatingState.eRun,     // 运行态 / Run state
    E_DL_CoatingState.eLimit:   // 限幅态 / Limit state
        bActive := TRUE;        // 闭环投入 / Loop active

        // ---- 测厚有效性：冻结积分、输出保持 / Invalid meas: freeze integral, hold output ----
        IF NOT bMeasValid THEN
            eErr    := 16#0002_371E;  // 信息级：测厚无效 / Info: meas invalid
            // fGapCmd_mm 保持不动（绝不因无测量而推进）/ Hold gap command
        ELSE
            // ---- 非有限测厚闸 / Non-finite measurement guard ----
            IF (fMeas_gsm <> fMeas_gsm) OR (ABS(fMeas_gsm) >= 1.0E12) THEN
                eErr := 16#0002_371E; // 按无效测厚处理 / Treat as invalid
            ELSE
                // ---- 一阶滤波（内联，alpha=0.2）/ Inline first-order filter ----
                fFilt_gsm := fFilt_gsm + 0.2 * (fMeas_gsm - fFilt_gsm);  // 一阶低通 / First-order LPF

                // ---- 新鲜偏差 / Fresh deviation ----
                fDevNow_gsm := fFilt_gsm - fSp_gsm;   // 偏差 / Deviation [g/m2]

                // ---- 死区判（防抖动磨模头）/ Dead band check ----
                fBandAbs := fSp_gsm * fBandPct / 100.0;  // 绝对带宽 / Absolute band [g/m2]
                IF ABS(fDevNow_gsm) <= fBandAbs THEN
                    bInBand := TRUE;    // 带内标志 / In-band flag
                    eErr    := 16#0002_371A;  // 信息级：带内不动作 / Info: in-band idle
                ELSE
                    // ---- 写入延时队列（循环缓冲）/ Write fresh deviation into delay queue ----
                    aDelayQ[uQHead] := fDevNow_gsm;   // 写入当前偏差 / Store fresh deviation
                    uQHead := uQHead + 1;             // 指针前移 / Advance pointer
                    IF uQHead >= uQLenCfg THEN
                        uQHead := 0;                  // 回绕 / Wrap around
                    END_IF
                    IF uQLen < uQLenCfg THEN
                        uQLen := uQLen + 1;           // 队列填充中 / Queue filling
                    END_IF

                    // ---- 读出滞后 tDeadTime 拍前的偏差 / Read delayed deviation ----
                    fDev_gsm := aDelayQ[uQHead];      // 滞后补偿后偏差 / Delayed deviation [g/m2]

                    // ---- 积分型无差调节：按增益换算间隙增量 / Integral-type adjustment ----
                    fRateStep := fRateMax_mm_s * tCycleS;  // 单拍速率步长 / Rate step per cycle [mm]
                    fTrimNew := fTrim_mm - fGain_mm_per_gsm * fDev_gsm;  // 目标修正 / Tentative trim [mm]

                    // ---- 增量限速 / Rate limiting ----
                    IF (fTrimNew - fTrim_mm) > fRateStep THEN
                        fTrimNew := fTrim_mm + fRateStep;  // 正向限速 / Positive slew limit
                    ELSIF (fTrimNew - fTrim_mm) < -fRateStep THEN
                        fTrimNew := fTrim_mm - fRateStep;  // 负向限速 / Negative slew limit
                    END_IF

                    // ---- 总量限幅 + 触限抗饱和 / Total clamp + anti-windup at limit ----
                    IF fTrimNew > fTrimMax_mm THEN
                        fTrimNew := fTrimMax_mm;   // 上限钳制 / Upper clamp
                        eState := E_DL_CoatingState.eLimit;  // 进入限幅态 / Enter limit state
                        eErr := 16#0002_371D;      // 信息级：触限 / Info: at limit
                    ELSIF fTrimNew < -fTrimMax_mm THEN
                        fTrimNew := -fTrimMax_mm;  // 下限钳制 / Lower clamp
                        eState := E_DL_CoatingState.eLimit;  // 进入限幅态 / Enter limit state
                        eErr := 16#0002_371D;      // 信息级：触限 / Info: at limit
                    ELSE
                        eErr := 16#0002_371A;      // 信息级：正常调节 / Info: normal
                    END_IF

                    // ---- 触限后停止同向积分：只在离限方向才更新 / Anti-windup: only move away from limit ----
                    IF (eState = E_DL_CoatingState.eLimit) AND (fTrim_mm = fTrimMax_mm) AND (fTrimNew > fTrim_mm) THEN
                        // 已在上限且继续同向：冻结 / At upper limit, same direction: freeze
                    ELSIF (eState = E_DL_CoatingState.eLimit) AND (fTrim_mm = -fTrimMax_mm) AND (fTrimNew < fTrim_mm) THEN
                        // 已在下限且继续同向：冻结 / At lower limit, same direction: freeze
                    ELSE
                        fTrim_mm := fTrimNew;      // 采纳修正 / Adopt trim
                    END_IF

                    // ---- 间隙命令 = 初始 + 修正 / Gap command = initial + trim ----
                    fGapCmd_mm := fGapInit_mm + fTrim_mm;  // 输出间隙命令 / Output gap command [mm]
                END_IF
            END_IF
        END_IF

        // ---- 限幅态回到运行态：修正脱离边界即回 eRun / Limit back to run when off boundary ----
        IF (eState = E_DL_CoatingState.eLimit)
           AND (ABS(fTrim_mm) < fTrimMax_mm) THEN
            eState := E_DL_CoatingState.eRun;  // 回运行态 / Back to run
        END_IF

    ELSE                        // 非法状态拦截 / Illegal state interception
        eState := E_DL_CoatingState.eFault;  // 落故障态 / Fall to fault
        bActive := FALSE;       // 闭环退出 / Loop inactive
        eErr := 16#0002_371B;   // 故障码 / Fault code
END_CASE

// ---- 使能撤销：冻结输出回空闲 / Disable: freeze and idle ----
IF NOT bEnable THEN
    bActive := FALSE;           // 闭环退出 / Loop inactive
    eState  := E_DL_CoatingState.eIdle;  // 回空闲 / Back to idle
END_IF

END_FUNCTION_BLOCK

(* ---- FB_DL_ControlOutputSlewWatch.st ---- *)
(*
  Name        : FB_DL_ControlOutputSlewWatch
  Category    : DL_Algo
  Version     : 1.0.1
  Purpose     : 控制输出变化率监视：逐拍算输出速率（%/s），判超速（超 fSlewMax）、爬行（推动但速率低于 fSlewCreep）、振荡（窗口内速率符号翻转次数超阈），供回路诊断定性；/ Watch control output slew rate: detect over-speed, creeping and oscillation via sign-flip count within a time-ordered window
  Changelog   : v1.0.1 R52 五抽终审修复首拍 _nHead=0 越界写（段1 域外自愈）
  Fix R54     : _nHead/_nFill 声明初值补齐（R52 五抽严重项），运行时自愈保留作双保险
  溯源        : 借 t2-1-lgf·measurement 的分类/参数域组织，clean-room 实现
  Boundary    : ① 扫描周期闸：tScan <= T#0S → 锁存故障（速率除零前置）；
                ② 符号翻转统计按时间序环回遍历（_nOldest→_nIdx，R52 环窗时间序范式），不做下标序直读；
                ③ 死区判据：|速率| <= eps 视为无方向（不参与符号翻转计数，防噪声刷计数）；
                ④ 窗口深度钳位 4..32，翻转阈 = 窗深 / 2（整数直比，无浮点）；
                ⑤ 全部判据为观测级，不写输出侧（属主边界：本件不动控制量）。
*)
TYPE E_DL_CswState :
(
    eIdle  := 0,                             (* 未使能 / Disabled *)
    eRun   := 10,                            (* 监视运行 / Watching *)
    eFault := 90                             (* 故障锁存相 / Fault latched *)
);
END_TYPE

TYPE E_DL_CswCause :
(
    eNone       := 0,                        (* 无故障成因 / No cause *)
    eCfgIllegal := 1,                        (* 组态非法：周期/速率阈值/窗深越域 / Illegal config *)
    ePhaseBad   := 2                         (* 非法相位兜底 / Illegal phase fallback *)
);
END_TYPE

FUNCTION_BLOCK FB_DL_ControlOutputSlewWatch
VAR_INPUT
    fOut       : REAL := 0.0;                (* 被监视控制输出（阀位/频率给定）[%] / Monitored control output *)
    tScan      : TIME := T#10MS;             (* 采样周期（速率除子），域 > T#0S [ms] / Sampling period, > 0 *)
    fSlewMax   : REAL := 50.0;               (* 允许速率上限，域 > 0 [%/s] / Allowed slew limit, > 0 *)
    fSlewCreep : REAL := 0.5;                (* 爬行判定下限（有效但过慢），域 0 < x < fSlewMax [%/s] / Creep lower limit *)
    nWinLen    : INT := 16;                  (* 符号翻转统计窗深，域 4..32 [点] / Flip window depth *)
    bEnable    : BOOL := TRUE;               (* 使能 [-] / Enable *)
    bReset     : BOOL := FALSE;              (* 复位命令，上升沿清窗口与全部标志 [-] / Reset command *)
END_VAR
VAR_OUTPUT
    fSlew      : REAL;                       (* 本拍输出速率 [%/s] / Output slew this scan *)
    fSlewPeak  : REAL;                       (* 窗口内 |速率| 峰值 [%/s] / Window peak absolute slew *)
    nFlips     : INT;                        (* 窗口内速率符号翻转次数 [-] / Sign flips within window *)
    bSlewHigh  : BOOL;                       (* 超速判据 [-] / Over-speed verdict *)
    bCreep     : BOOL;                       (* 爬行判据 [-] / Creeping verdict *)
    bOscillate : BOOL;                       (* 振荡判据（翻转次数超半窗）[-] / Oscillation verdict *)
    eState     : E_DL_CswState;              (* 状态出口 / State outlet *)
    eCause     : E_DL_CswCause;              (* 故障成因出口（R190 归因唯一） / Fault cause outlet *)
    bError     : BOOL;                       (* 故障锁存标志 [-] / Fault latch flag *)
END_VAR
VAR
    _eState  : E_DL_CswState := E_DL_CswState.eIdle;     (* 内部相位（CASE 唯一写入目标） / Internal phase *)
    _eCause  : E_DL_CswCause := E_DL_CswCause.eNone;     (* 故障成因锁存量 / Latched cause *)
    rtReset  : R_TRIG;                       (* 复位沿实例，段 0 无条件调用 / Reset edge instance *)
    _bFault  : BOOL;                         (* 故障锁存位 / Latched fault bit *)
    _bCfgBad : BOOL;                         (* 组态非法当拍量 / Illegal config this scan *)
    _bInit   : BOOL;                         (* 前值初始化标志（首拍速率按 0） / First-scan init *)
    _fPrev   : REAL;                         (* 上拍输出快照 [%] / Previous output snapshot *)
    _fDtSec  : REAL;                         (* 周期折算秒值，域 > eps [s] / Period in seconds *)
    _fPeak   : REAL;                         (* 窗口峰值累加量 [%/s] / Peak accumulator *)
    _aSign   : ARRAY[1..32] OF INT;          (* 速率符号环窗（-1/0/+1）[-] / Slew sign ring window *)
    _nHead   : INT := 1;                     (* 环形写入头游标（声明期安全初值，R194）[-] / Ring head cursor, declared init *)
    _nFill   : INT := 0;                     (* 窗口填充数（声明期安全初值，R194）[点] / Fill count, declared init *)
    _nEff    : INT;                          (* 钳位后生效窗深 [点] / Clamped depth *)
    _nOldest : INT;                          (* 最旧样本槽位（每趟重算）[-] / Oldest slot *)
    _nIdx    : INT;                          (* 时间序 → 环形槽位换算下标 [-] / Time-order to slot index *)
    _nJ      : INT;                          (* 时间序游标 0.._nFill-1 [-] / Time cursor *)
    _nFlip   : INT;                          (* 翻转计数累加量 [-] / Flip accumulator *)
    _nPrevSg : INT;                          (* 上一非零符号（时间序传播）[-] / Previous non-zero sign *)
    _nSg     : INT;                          (* 本点符号 [-] / Sign of current point *)
    _nFlipThr: INT;                          (* 翻转阈值 = 窗深 / 2 [-] / Flip threshold *)
END_VAR
VAR CONSTANT
    DL_CSW_EPS    : REAL := 1.0E-6;          (* 速率死区判零容差 [%/s] / Slew deadband epsilon *)
    DL_CSW_NMAX   : INT  := 32;              (* 窗深容量上限 [点] / Window capacity limit *)
    DL_CSW_NMIN   : INT  := 4;               (* 窗深下限 [点] / Window depth lower bound *)
    DL_CSW_SG_P   : INT  := 1;               (* 正符号编码 [-] / Positive sign code *)
    DL_CSW_SG_N   : INT  := -1;              (* 负符号编码 [-] / Negative sign code *)
    DL_CSW_SG_Z   : INT  := 0;               (* 零符号编码（无方向，不参与翻转）[-] / Zero sign code *)
END_VAR

(* —— 段 0：当拍判据派生 + 实例无条件刷新（R228A） —— *)
_fDtSec := TIME_TO_LREAL(tScan) / 1000.0;                                      (* 周期秒化（除子常量 1000） / Period to seconds *)
_bCfgBad := NOT (tScan > T#0S)                                                 (* 周期正域闸 / Period gate *)
            OR (fSlewMax <= DL_CSW_EPS)                                        (* 速率上限正域闸 / Slew limit gate *)
            OR (fSlewCreep < 0.0) OR (fSlewCreep >= fSlewMax)                  (* 爬行下限域闸 0 <= x < max / Creep gate *)
            OR (nWinLen < DL_CSW_NMIN) OR (nWinLen > DL_CSW_NMAX);             (* 窗深域闸（也保证翻转统计有界） / Depth gate *)
rtReset(CLK := bReset);                                                        (* 复位沿每拍必调 / Reset edge every scan *)
_nEff := nWinLen;                                                              (* 生效窗深初值 / Depth init *)
IF _nEff < DL_CSW_NMIN THEN
    _nEff := DL_CSW_NMIN;                                                      (* 下限钳位 / Lower clamp *)
END_IF
IF _nEff > DL_CSW_NMAX THEN
    _nEff := DL_CSW_NMAX;                                                      (* 上限钳位（R308） / Upper clamp *)
END_IF
IF _nEff < 2 THEN
    _nEff := 2;                                                                (* 兜底防除零（阈计算分母） / Fallback guard *)
END_IF
_nFlipThr := _nEff / 2;                                                        (* 翻转阈值（整数除，分母 >= 2） / Flip threshold *)

(* —— 段 1：单拍量预清零（R107） —— *)
bSlewHigh := FALSE;                                                            (* 超速判据预清 / Over-speed preset *)
bCreep := FALSE;                                                               (* 爬行判据预清 / Creep preset *)
bOscillate := FALSE;                                                           (* 振荡判据预清 / Oscillation preset *)
nFlips := 0;                                                                   (* 翻转数预清 / Flip count preset *)
fSlew := 0.0;                                                                  (* 速率预清（首拍/失能路径） / Slew preset *)
IF (_nHead < 1) OR (_nHead > _nEff) THEN
    _nHead := 1;                                                               (* 头游标域外自愈：首拍 0 与窗深缩小后回钳（v1.0.1） / Head self-heal *)
END_IF
IF _nFill > _nEff THEN
    _nFill := _nEff;                                                           (* 填充数随窗深回钳 / Fill clamped to depth *)
END_IF

(* —— 段 2：复位沿处理（作用域：清故障 + 清窗 + 清峰值 + 迁 eIdle，R283 逐项声明） —— *)
IF rtReset.Q THEN
    _bFault := FALSE;                                                          (* 清故障锁存 / Clear fault *)
    _eCause := E_DL_CswCause.eNone;                                            (* 清成因 / Clear cause *)
    _nFill := 0;                                                               (* 清窗填充 / Clear fill *)
    _nHead := 1;                                                               (* 头游标复位 / Head reset *)
    _nOldest := 1;                                                             (* 最旧槽复位 / Oldest reset *)
    _fPeak := 0.0;                                                             (* 清峰值 / Clear peak *)
    _fPrev := 0.0;                                                             (* 清前值 / Clear previous *)
    _bInit := FALSE;                                                           (* 清初始化标志 / Clear init *)
    fSlewPeak := 0.0;                                                          (* 清峰值出口 / Clear peak outlet *)
    _eState := E_DL_CswState.eIdle;                                            (* 迁未使能相 / Back to idle *)
END_IF

(* —— 段 3：组态故障锁存（锁存至复位沿，R189） —— *)
IF _bCfgBad AND NOT _bFault THEN
    _bFault := TRUE;                                                           (* 锁存故障位 / Latch fault *)
    _eCause := E_DL_CswCause.eCfgIllegal;                                      (* 成因：组态非法 / Cause: illegal config *)
    _eState := E_DL_CswState.eFault;                                           (* 同步迁故障相 / Migrate to fault *)
END_IF

(* —— 段 4：CASE 主状态机（ELSE 兜底迁 eFault，红线 6） —— *)
CASE _eState OF
    E_DL_CswState.eIdle:                                                       (* 未使能：不采集，出口保持 0 / Disabled *)
        _bInit := FALSE;                                                       (* 失能清初始化（重使能重新对齐） / Clear init *)
        IF bEnable AND NOT _bFault THEN
            _eState := E_DL_CswState.eRun;                                     (* 使能进入监视 / Enter watching *)
        END_IF
    E_DL_CswState.eRun:                                                        (* 监视相：速率 + 符号窗 + 三判据 / Watching *)
        IF NOT bEnable THEN
            _eState := E_DL_CswState.eIdle;                                    (* 失能回未使能 / Back to idle *)
        ELSIF (_fDtSec > DL_CSW_EPS) THEN
            IF NOT _bInit THEN
                _fPrev := fOut;                                                (* 首拍对齐：速率按 0，不产虚假尖峰 / First-scan alignment *)
                _bInit := TRUE;                                                (* 立初始化标志 / Set init *)
            END_IF
            fSlew := (fOut - _fPrev) / _fDtSec;                                (* 输出速率：除子已过闸 [%/s] / Slew, divisor gated *)
            _fPrev := fOut;                                                    (* 快照推进 / Advance snapshot *)
            IF fSlew > DL_CSW_EPS THEN
                _nSg := DL_CSW_SG_P;                                           (* 正方向 / Rising *)
            ELSIF fSlew < (-DL_CSW_EPS) THEN
                _nSg := DL_CSW_SG_N;                                           (* 负方向 / Falling *)
            ELSE
                _nSg := DL_CSW_SG_Z;                                           (* 带内：无方向（不参与翻转） / Deadband: no direction *)
            END_IF
            _aSign[_nHead] := _nSg;                                            (* 符号入环窗（下标已 1.._nEff 钳位） / Sign into ring *)
            _nHead := _nHead + 1;                                              (* 头游标递进 / Head advance *)
            IF _nHead > _nEff THEN
                _nHead := 1;                                                   (* 环回卷 / Ring wrap *)
            END_IF
            IF _nFill < _nEff THEN
                _nFill := _nFill + 1;                                          (* 填充封顶 / Fill cap *)
            END_IF
            IF _nFill >= 1 THEN
                _nOldest := _nHead - _nFill;                                   (* 最旧槽：未满窗 = 1 / Oldest while filling *)
                IF _nOldest < 1 THEN
                    _nOldest := _nOldest + _nEff;                              (* 满窗回卷：最旧在 _nHead 槽（R52 时间序） / Wrapped oldest *)
                END_IF
            END_IF
            _nFlip := 0;                                                       (* 翻转计数每趟重置（R227） / Flips reset per pass *)
            _nPrevSg := DL_CSW_SG_Z;                                           (* 前符号预置为零（时间序起点） / Previous sign preset *)
            _fPeak := 0.0;                                                     (* 峰值每趟重算 / Peak recompute *)
            _nJ := 0;                                                          (* 时间序游标起头 / Time cursor reset *)
            WHILE _nJ < _nFill DO                                              (* 按时间序环回遍历（R52 范式） / Time-ordered ring walk *)
                _nIdx := _nOldest + _nJ;                                       (* 时间序 → 槽位映射 / Time order to slot *)
                IF _nIdx > _nEff THEN
                    _nIdx := _nIdx - _nEff;                                    (* 槽位环回 / Slot wrap *)
                END_IF
                _nSg := _aSign[_nIdx];                                         (* 该点符号 / Sign of point *)
                IF _nSg <> DL_CSW_SG_Z THEN
                    IF (_nPrevSg <> DL_CSW_SG_Z) AND (_nSg <> _nPrevSg) THEN
                        _nFlip := _nFlip + 1;                                  (* 非零符号相反：计一次翻转 / Opposite non-zero signs *)
                    END_IF
                    _nPrevSg := _nSg;                                          (* 有效符号向前传播 / Propagate last valid sign *)
                END_IF
                _nJ := _nJ + 1;                                                (* 游标递进 / Cursor advance *)
            END_WHILE
            nFlips := _nFlip;                                                  (* 翻转数出口 / Flip outlet *)
            IF ABS(fSlew) > _fPeak THEN
                _fPeak := ABS(fSlew);                                          (* 本拍更新窗口 |速率| 峰值 / Update peak *)
            END_IF
            fSlewPeak := _fPeak;                                               (* 峰值出口 / Peak outlet *)
            IF ABS(fSlew) > fSlewMax THEN
                bSlewHigh := TRUE;                                             (* 超速判据（ABS 差比较，禁单侧） / Over-speed verdict *)
            END_IF
            IF (ABS(fSlew) > DL_CSW_EPS) AND (ABS(fSlew) < fSlewCreep) THEN
                bCreep := TRUE;                                                (* 爬行判据：动了但过慢 / Creeping verdict *)
            END_IF
            IF _nFlip >= _nFlipThr THEN
                bOscillate := TRUE;                                            (* 振荡判据：翻转过半窗 / Oscillation verdict *)
            END_IF
        END_IF
    E_DL_CswState.eFault:                                                      (* 故障相：冻结保持末值，仅复位沿出 / Fault *)
        ;                                                                      (* 锁存回放（R28） / Replay from latch *)
    ELSE                                                                       (* 非法相位兜底迁安全态 / Illegal phase fallback *)
        _eState := E_DL_CswState.eFault;                                       (* 迁故障相 / To fault *)
        _bFault := TRUE;                                                       (* 同步锁存 / Latch *)
        _eCause := E_DL_CswCause.ePhaseBad;                                    (* 成因：非法相位 / Cause: illegal phase *)
END_CASE

(* —— 段 5：出口映射（bError/eState 同源，R191） —— *)
bError := _bFault;                                                             (* 故障标志镜像 / Fault flag mirror *)
eState := _eState;                                                             (* 状态出口 / State outlet *)
eCause := _eCause;                                                             (* 成因出口 / Cause outlet *)
END_FUNCTION_BLOCK
